(* IEC 61131-3 sources: deprecated-refusr-repo/GP/Main/samples (part 24) *)

(* ---- RND-EXPR_trial-nosed-gunky.st ---- *)
(*
This code implements a randomly grown symbolic expression:

(!(IN26 & (IN45 | ((xor(xor(IN3, !(xor(xor((IN43 & IN34) | (IN19 | IN26), xor(xor(!(IN50), IN21 | IN1), IN17 & IN23)), xor(xor(xor(xor(IN4, IN2), IN41), IN7 & IN29), IN13)))), IN42)) | IN20)))) | (!((xor(xor(!(!(xor(xor(!((!(IN14)) & IN36), ((xor(xor(IN45, IN34), IN41)) | (IN17 | IN11)) & IN16), !(xor(xor(IN37 & IN25, true), IN17 & IN22))))), !((!(IN31)) | (!(IN6)))), ((!(IN16)) | IN27) & (IN46 & ((xor(xor(!(IN15 | IN34), IN28), !(IN7 & IN3))) & ((xor(xor(!(IN32), xor(xor(IN36, IN43), IN28)), !(IN36))) & IN44))))) & IN13))

*)

FUNCTION_BLOCK F_CollectInput
  VAR_IN_OUT
      Data : ARRAY[1..50] OF BOOL;
  END_VAR
  VAR_INPUT
      TICK  : BOOL := 0;
      IN1   : BOOL := 0;
      IN2   : BOOL := 0;
      IN3   : BOOL := 0;
      IN4   : BOOL := 0;
      IN5   : BOOL := 0;
      RESET : BOOL := FALSE;
  END_VAR
  VAR_OUTPUT
      Finished : BOOL;
  END_VAR
  VAR
      j    : USINT := 1;
      tock : BOOL  := 0;
  END_VAR
  IF NOT RESET AND tock = NOT TICK THEN
      Data[j]   := IN1;
      Data[j+1] := IN2;
      Data[j+2] := IN3;
      Data[j+3] := IN4;
      Data[j+4] := IN5;
      j := j + 5;
      tock := TICK;
  ELSE
      j := 1;
      tock := 0;
  END_IF;
  Finished := (j > 50);
END_FUNCTION_BLOCK

PROGRAM Boiler
  VAR
    Data  : ARRAY[1..50] OF BOOL;
    Ready : BOOL;
    CollectInput : F_CollectInput;
  END_VAR
  VAR
    TICK     AT %IX1.0 : BOOL;
    IN1      AT %IX0.3 : BOOL;
    IN2      AT %IX0.4 : BOOL;
    IN3      AT %IX0.5 : BOOL;
    IN4      AT %IX0.6 : BOOL;
    IN5      AT %IX0.7 : BOOL;
    OutReady AT %QX0.0 : BOOL := FALSE;
    FeedNext AT %QX0.1 : BOOL := FALSE;
    Out      AT %QX0.2 : BOOL;
  END_VAR
  CollectInput(TICK:=TICK, IN1:=IN1, IN2:=IN2, IN3:=IN3, IN4:=IN4, IN5:=IN5);
  Ready := CollectInput.Finished;
  FeedNext := 1;
  IF Ready THEN
    Out := ((NOT (Data[26] AND (Data[45] OR (((Data[3] XOR (NOT ((((Data[43] AND Data[34]) OR (Data[19] OR Data[26])) XOR (((NOT Data[50]) XOR (Data[21] OR Data[1])) XOR (Data[17] AND Data[23]))) XOR ((((Data[4] XOR Data[2]) XOR Data[41]) XOR (Data[7] AND Data[29])) XOR Data[13])))) XOR Data[42]) OR Data[20])))) OR (NOT ((((NOT (NOT (((NOT ((NOT Data[14]) AND Data[36])) XOR ((((Data[45] XOR Data[34]) XOR Data[41]) OR (Data[17] OR Data[11])) AND Data[16])) XOR (NOT (((Data[37] AND Data[25]) XOR TRUE) XOR (Data[17] AND Data[22])))))) XOR (NOT ((NOT Data[31]) OR (NOT Data[6])))) XOR (((NOT Data[16]) OR Data[27]) AND (Data[46] AND ((((NOT (Data[15] OR Data[34])) XOR Data[28]) XOR (NOT (Data[7] AND Data[3]))) AND ((((NOT Data[32]) XOR ((Data[36] XOR Data[43]) XOR Data[28])) XOR (NOT Data[36])) AND Data[44]))))) AND Data[13])));
    OutReady := 1;
    CollectInput(RESET:=TRUE);
  END_IF;
END_PROGRAM

CONFIGURATION Config0
  RESOURCE Res0 ON PLC
    TASK task0(INTERVAL := T#20ms,PRIORITY := 0);
    PROGRAM instance0 WITH task0 : Boiler;
  END_RESOURCE
END_CONFIGURATION

(* ---- RND-EXPR_trill-blare-frail.st ---- *)
(*
This code implements a randomly grown symbolic expression:

(xor(xor(xor(xor((((((xor(xor(!(IN12), !(IN17)), xor(xor(IN9, IN18), IN16))) | (!(!(IN37)))) | IN16) & (xor(xor(IN45, (xor(xor(IN41 | IN9, xor(xor(IN35, IN31), IN31)), false & IN31)) | ((xor(xor(IN20, IN44), IN36)) | (IN7 & IN36))), false & IN37))) | IN2) | (IN40 & (xor(xor((xor(xor(xor(xor(IN13, IN26), IN49 | IN33), (xor(xor(IN9, IN4), IN10)) & IN35), (xor(xor(IN38, IN22), IN49)) & (IN26 | IN2))) & (xor(xor((IN21 | IN37) | IN35, xor(xor(xor(xor(IN27, IN35), IN49), IN20), !(IN38))), xor(xor(!(IN24), IN47 & IN9), IN49 & IN17))), (IN2 & ((xor(xor(IN39, true), IN43)) | (!(IN6)))) & (xor(xor(xor(xor(IN32 | IN28, !(IN19)), IN40 | IN22), !(IN3 & IN26)), (IN29 | IN25) | (IN45 & IN27)))), xor(xor((!(IN44)) & IN6, IN29), (!(IN7 & IN11)) | ((false & IN15) | (!(IN19))))))), IN17), xor(xor((IN38 & (IN15 | ((IN27 | (!(IN8))) & (IN23 | (IN11 & IN7))))) | (xor(xor((((xor(xor(IN34, IN2), IN40)) | IN1) | (!(IN9 | IN21))) & (!(xor(xor(IN30 | IN29, xor(xor(IN44, IN42), IN31)), true & IN38))), (IN10 | ((IN10 | IN13) & (IN25 | IN48))) & IN18), xor(xor(!(xor(xor(!(IN15), IN14 & IN49), false)), IN16), IN33))), IN13), xor(xor(!((((!(IN21)) & IN46) | (!(!(IN30)))) | (!((xor(xor(IN29, IN30), IN17)) | (xor(xor(IN48, IN6), IN1))))), xor(xor(!(IN18), (((!(IN34)) & (IN25 | IN49)) & (!(IN46 | IN49))) & (!(xor(xor(xor(xor(IN12, IN43), IN16), IN41), IN17)))), IN11 | (IN5 | false))), ((((!(IN35)) | (xor(xor(IN23, IN39), IN8))) & IN6) & (!(xor(xor(IN21 & IN34, true | IN14), xor(xor(IN23, IN26), IN5))))) & IN28))), !(!(IN4))), (IN38 | (xor(xor(!(IN16 | (IN25 & (!(!(IN31))))), xor(xor(xor(xor((false | (xor(xor(IN33, IN12), IN48))) | ((xor(xor(IN5, IN49), IN14)) & IN11), !((IN49 | IN29) | (IN29 & IN12))), ((IN48 | IN19) | (IN10 | IN4)) | ((!(IN37)) & (IN39 & IN4))), (!((IN33 | true) | (xor(xor(IN26, IN44), IN22)))) | (IN37 | (xor(xor(IN30 | IN33, IN47), !(IN7))))), (!(xor(xor(!(IN21), !(IN11)), !(IN17)))) & IN12)), xor(xor((((!(IN22)) | (IN18 & IN6)) & (xor(xor(xor(xor(IN30, IN18), IN11), IN14 & IN13), IN18 & IN44))) & (xor(xor(IN30 & (IN31 & IN44), xor(xor(xor(xor(IN22, IN16), IN17), xor(xor(IN13, IN42), IN23)), IN38 & IN3)), !(xor(xor(IN41, IN47), IN26)))), IN3), IN12 | IN1)))) & (xor(xor(IN30, !(xor(xor(xor(xor(IN49 & (!(!(IN12))), IN12 & (!(IN13 | IN31))), !((IN21 | IN45) & (IN43 | IN21))), xor(xor(!((IN24 | IN34) | (!(IN1))), ((!(IN44)) & (xor(xor(IN20, IN30), IN17))) | (xor(xor(IN23 & IN49, IN45 & IN25), !(IN34)))), !((!(IN13)) | (xor(xor(IN49, IN15), IN41))))), ((IN4 & (IN19 & IN39)) | ((xor(xor(IN9, IN46), IN40)) & (IN30 & IN45))) & (IN49 | IN13)))), xor(xor(xor(xor(((IN50 & (!(IN24))) & ((IN47 | IN39) & (IN40 & IN24))) & ((xor(xor(IN10 | IN23, IN7 | IN31), IN15 | IN34)) & (IN44 | (!(IN46)))), !(xor(xor(xor(xor(IN29, IN20), IN41 & IN28), IN12), IN27 & (xor(xor(IN42, IN24), IN2))))), IN23), IN11), ((((xor(xor(IN44, IN30), IN46)) | IN35) & IN44) | ((IN45 | (IN7 | IN9)) & IN40)) & IN26))))) | (!((((((xor(xor(IN40, xor(xor(IN25 & IN33, !(IN30)), xor(xor(IN17, IN41), IN29))), IN23)) | (!(xor(xor(xor(xor(IN16, IN49), IN38), IN2 | IN47), IN6 | IN24)))) | IN9) | (!(IN10))) | IN25) & (IN47 | (!(((!(!(IN41 & IN48))) | (IN6 | IN11)) & (((IN12 & IN38) & IN8) | ((xor(xor(IN39 & IN14, IN34 | IN30), xor(xor(IN23, IN46), IN33))) | IN49)))))))

*)

FUNCTION_BLOCK F_CollectInput
  VAR_IN_OUT
      Data : ARRAY[1..50] OF BOOL;
  END_VAR
  VAR_INPUT
      TICK  : BOOL := 0;
      IN1   : BOOL := 0;
      IN2   : BOOL := 0;
      IN3   : BOOL := 0;
      IN4   : BOOL := 0;
      IN5   : BOOL := 0;
      RESET : BOOL := FALSE;
  END_VAR
  VAR_OUTPUT
      Finished : BOOL;
  END_VAR
  VAR
      j    : USINT := 1;
      tock : BOOL  := 0;
  END_VAR
  IF NOT RESET AND tock = NOT TICK THEN
      Data[j]   := IN1;
      Data[j+1] := IN2;
      Data[j+2] := IN3;
      Data[j+3] := IN4;
      Data[j+4] := IN5;
      j := j + 5;
      tock := TICK;
  ELSE
      j := 1;
      tock := 0;
  END_IF;
  Finished := (j > 50);
END_FUNCTION_BLOCK

PROGRAM Boiler
  VAR
    Data  : ARRAY[1..50] OF BOOL;
    Ready : BOOL;
    CollectInput : F_CollectInput;
  END_VAR
  VAR
    TICK     AT %IX1.0 : BOOL;
    IN1      AT %IX0.3 : BOOL;
    IN2      AT %IX0.4 : BOOL;
    IN3      AT %IX0.5 : BOOL;
    IN4      AT %IX0.6 : BOOL;
    IN5      AT %IX0.7 : BOOL;
    OutReady AT %QX0.0 : BOOL := FALSE;
    FeedNext AT %QX0.1 : BOOL := FALSE;
    Out      AT %QX0.2 : BOOL;
  END_VAR
  CollectInput(TICK:=TICK, IN1:=IN1, IN2:=IN2, IN3:=IN3, IN4:=IN4, IN5:=IN5);
  Ready := CollectInput.Finished;
  FeedNext := 1;
  IF Ready THEN
    Out := (((((((((((((NOT Data[12]) XOR (NOT Data[17])) XOR ((Data[9] XOR Data[18]) XOR Data[16])) OR (NOT (NOT Data[37]))) OR Data[16]) AND ((Data[45] XOR ((((Data[41] OR Data[9]) XOR ((Data[35] XOR Data[31]) XOR Data[31])) XOR (FALSE AND Data[31])) OR (((Data[20] XOR Data[44]) XOR Data[36]) OR (Data[7] AND Data[36])))) XOR (FALSE AND Data[37]))) OR Data[2]) OR (Data[40] AND (((((((Data[13] XOR Data[26]) XOR (Data[49] OR Data[33])) XOR (((Data[9] XOR Data[4]) XOR Data[10]) AND Data[35])) XOR (((Data[38] XOR Data[22]) XOR Data[49]) AND (Data[26] OR Data[2]))) AND ((((Data[21] OR Data[37]) OR Data[35]) XOR ((((Data[27] XOR Data[35]) XOR Data[49]) XOR Data[20]) XOR (NOT Data[38]))) XOR (((NOT Data[24]) XOR (Data[47] AND Data[9])) XOR (Data[49] AND Data[17])))) XOR ((Data[2] AND (((Data[39] XOR TRUE) XOR Data[43]) OR (NOT Data[6]))) AND (((((Data[32] OR Data[28]) XOR (NOT Data[19])) XOR (Data[40] OR Data[22])) XOR (NOT (Data[3] AND Data[26]))) XOR ((Data[29] OR Data[25]) OR (Data[45] AND Data[27]))))) XOR ((((NOT Data[44]) AND Data[6]) XOR Data[29]) XOR ((NOT (Data[7] AND Data[11])) OR ((FALSE AND Data[15]) OR (NOT Data[19]))))))) XOR Data[17]) XOR ((((Data[38] AND (Data[15] OR ((Data[27] OR (NOT Data[8])) AND (Data[23] OR (Data[11] AND Data[7]))))) OR (((((((Data[34] XOR Data[2]) XOR Data[40]) OR Data[1]) OR (NOT (Data[9] OR Data[21]))) AND (NOT (((Data[30] OR Data[29]) XOR ((Data[44] XOR Data[42]) XOR Data[31])) XOR (TRUE AND Data[38])))) XOR ((Data[10] OR ((Data[10] OR Data[13]) AND (Data[25] OR Data[48]))) AND Data[18])) XOR (((NOT (((NOT Data[15]) XOR (Data[14] AND Data[49])) XOR FALSE)) XOR Data[16]) XOR Data[33]))) XOR Data[13]) XOR (((NOT ((((NOT Data[21]) AND Data[46]) OR (NOT (NOT Data[30]))) OR (NOT (((Data[29] XOR Data[30]) XOR Data[17]) OR ((Data[48] XOR Data[6]) XOR Data[1]))))) XOR (((NOT Data[18]) XOR ((((NOT Data[34]) AND (Data[25] OR Data[49])) AND (NOT (Data[46] OR Data[49]))) AND (NOT ((((Data[12] XOR Data[43]) XOR Data[16]) XOR Data[41]) XOR Data[17])))) XOR (Data[11] OR (Data[5] OR FALSE)))) XOR (((((NOT Data[35]) OR ((Data[23] XOR Data[39]) XOR Data[8])) AND Data[6]) AND (NOT (((Data[21] AND Data[34]) XOR (TRUE OR Data[14])) XOR ((Data[23] XOR Data[26]) XOR Data[5])))) AND Data[28])))) XOR (NOT (NOT Data[4]))) XOR ((Data[38] OR (((NOT (Data[16] OR (Data[25] AND (NOT (NOT Data[31]))))) XOR ((((((FALSE OR ((Data[33] XOR Data[12]) XOR Data[48])) OR (((Data[5] XOR Data[49]) XOR Data[14]) AND Data[11])) XOR (NOT ((Data[49] OR Data[29]) OR (Data[29] AND Data[12])))) XOR (((Data[48] OR Data[19]) OR (Data[10] OR Data[4])) OR ((NOT Data[37]) AND (Data[39] AND Data[4])))) XOR ((NOT ((Data[33] OR TRUE) OR ((Data[26] XOR Data[44]) XOR Data[22]))) OR (Data[37] OR (((Data[30] OR Data[33]) XOR Data[47]) XOR (NOT Data[7]))))) XOR ((NOT (((NOT Data[21]) XOR (NOT Data[11])) XOR (NOT Data[17]))) AND Data[12]))) XOR ((((((NOT Data[22]) OR (Data[18] AND Data[6])) AND ((((Data[30] XOR Data[18]) XOR Data[11]) XOR (Data[14] AND Data[13])) XOR (Data[18] AND Data[44]))) AND (((Data[30] AND (Data[31] AND Data[44])) XOR ((((Data[22] XOR Data[16]) XOR Data[17]) XOR ((Data[13] XOR Data[42]) XOR Data[23])) XOR (Data[38] AND Data[3]))) XOR (NOT ((Data[41] XOR Data[47]) XOR Data[26])))) XOR Data[3]) XOR (Data[12] OR Data[1])))) AND ((Data[30] XOR (NOT (((((Data[49] AND (NOT (NOT Data[12]))) XOR (Data[12] AND (NOT (Data[13] OR Data[31])))) XOR (NOT ((Data[21] OR Data[45]) AND (Data[43] OR Data[21])))) XOR (((NOT ((Data[24] OR Data[34]) OR (NOT Data[1]))) XOR (((NOT Data[44]) AND ((Data[20] XOR Data[30]) XOR Data[17])) OR (((Data[23] AND Data[49]) XOR (Data[45] AND Data[25])) XOR (NOT Data[34])))) XOR (NOT ((NOT Data[13]) OR ((Data[49] XOR Data[15]) XOR Data[41]))))) XOR (((Data[4] AND (Data[19] AND Data[39])) OR (((Data[9] XOR Data[46]) XOR Data[40]) AND (Data[30] AND Data[45]))) AND (Data[49] OR Data[13]))))) XOR (((((((Data[50] AND (NOT Data[24])) AND ((Data[47] OR Data[39]) AND (Data[40] AND Data[24]))) AND ((((Data[10] OR Data[23]) XOR (Data[7] OR Data[31])) XOR (Data[15] OR Data[34])) AND (Data[44] OR (NOT Data[46])))) XOR (NOT ((((Data[29] XOR Data[20]) XOR (Data[41] AND Data[28])) XOR Data[12]) XOR (Data[27] AND ((Data[42] XOR Data[24]) XOR Data[2]))))) XOR Data[23]) XOR Data[11]) XOR ((((((Data[44] XOR Data[30]) XOR Data[46]) OR Data[35]) AND Data[44]) OR ((Data[45] OR (Data[7] OR Data[9])) AND Data[40])) AND Data[26]))))) OR (NOT (((((((Data[40] XOR (((Data[25] AND Data[33]) XOR (NOT Data[30])) XOR ((Data[17] XOR Data[41]) XOR Data[29]))) XOR Data[23]) OR (NOT ((((Data[16] XOR Data[49]) XOR Data[38]) XOR (Data[2] OR Data[47])) XOR (Data[6] OR Data[24])))) OR Data[9]) OR (NOT Data[10])) OR Data[25]) AND (Data[47] OR (NOT (((NOT (NOT (Data[41] AND Data[48]))) OR (Data[6] OR Data[11])) AND (((Data[12] AND Data[38]) AND Data[8]) OR ((((Data[39] AND Data[14]) XOR (Data[34] OR Data[30])) XOR ((Data[23] XOR Data[46]) XOR Data[33])) OR Data[49]))))))));
    OutReady := 1;
    CollectInput(RESET:=TRUE);
  END_IF;
END_PROGRAM

CONFIGURATION Config0
  RESOURCE Res0 ON PLC
    TASK task0(INTERVAL := T#20ms,PRIORITY := 0);
    PROGRAM instance0 WITH task0 : Boiler;
  END_RESOURCE
END_CONFIGURATION

(* ---- RND-EXPR_tulle-bench-aloha.st ---- *)
(*
This code implements a randomly grown symbolic expression:

(IN29 | (((!(IN27)) | (xor(xor(!(xor(xor(!((!(IN8)) & IN9), xor(xor(xor(xor(xor(xor(IN14, IN9), IN41), xor(xor(IN8, IN28), false)), xor(xor(IN9, IN9), IN2)), !(xor(xor(IN2, IN5), IN41))), (!(IN28)) & (xor(xor(IN12, IN39), IN7)))), IN36)), xor(xor(true, !(((IN30 | IN20) | IN9) & IN3)), xor(xor(false, (!(IN31)) | (xor(xor(IN41 | IN5, IN49 & IN1), !(IN13)))), xor(xor((IN28 | IN50) | (!(IN16)), (xor(xor(IN42, IN4), IN6)) | (xor(xor(IN38, IN42), IN36))), (xor(xor(IN46, IN18), IN35)) & (IN39 & IN11))))), IN39))) & (!(xor(xor(IN22 | ((!(xor(xor(IN21, IN5), IN41 & IN1))) | (xor(xor(xor(xor(IN15 | IN13, IN38 | IN6), !(IN1)), IN29), IN48))), IN18), IN3))))) | (!(!((((IN22 | (xor(xor(!(xor(xor(IN30, false), IN5)), !(IN14 | IN3)), !(IN48)))) | ((((!(IN28)) & (xor(xor(IN29, IN6), IN15))) & ((IN8 & IN49) | IN23)) & (((IN12 & IN1) | (xor(xor(IN43, IN5), IN47))) & ((!(IN33)) | (true | IN20))))) & ((!(IN50 | (!(IN5 | IN30)))) & IN40)) & (xor(xor((xor(xor((xor(xor(xor(xor(IN22, IN30), IN10), IN50), IN23 | IN47)) | (IN1 & (xor(xor(IN46, IN29), IN24))), IN24), ((IN2 & IN18) | (IN26 | IN47)) | ((!(IN19)) & IN35))) | ((IN33 & (!(IN25 | IN20))) | (xor(xor((xor(xor(IN40, IN13), IN19)) & (xor(xor(IN2, IN37), IN10)), (IN49 | IN40) & IN19), (xor(xor(IN25, IN24), IN14)) & (IN22 & IN32)))), (!(!((xor(xor(IN42, IN8), IN1)) & (!(IN42))))) & ((!(IN23 & IN19)) | ((!(IN29 & IN50)) & (!(IN8 & IN35))))), !(xor(xor(xor(xor((IN29 & IN22) & (!(IN14)), (IN32 & IN20) & (xor(xor(IN7, IN24), IN7))), (true & IN45) | (IN31 | IN44)), (xor(xor(!(IN45), IN35 | IN9), IN40 | IN3)) | ((xor(xor(IN5, IN37), IN27)) | (xor(xor(IN25, IN45), IN32)))), (false & (IN9 | IN18)) | (xor(xor(IN8, xor(xor(IN10, IN26), IN25)), !(IN39))))))))))

*)

FUNCTION_BLOCK F_CollectInput
  VAR_IN_OUT
      Data : ARRAY[1..50] OF BOOL;
  END_VAR
  VAR_INPUT
      TICK  : BOOL := 0;
      IN1   : BOOL := 0;
      IN2   : BOOL := 0;
      IN3   : BOOL := 0;
      IN4   : BOOL := 0;
      IN5   : BOOL := 0;
      RESET : BOOL := FALSE;
  END_VAR
  VAR_OUTPUT
      Finished : BOOL;
  END_VAR
  VAR
      j    : USINT := 1;
      tock : BOOL  := 0;
  END_VAR
  IF NOT RESET AND tock = NOT TICK THEN
      Data[j]   := IN1;
      Data[j+1] := IN2;
      Data[j+2] := IN3;
      Data[j+3] := IN4;
      Data[j+4] := IN5;
      j := j + 5;
      tock := TICK;
  ELSE
      j := 1;
      tock := 0;
  END_IF;
  Finished := (j > 50);
END_FUNCTION_BLOCK

PROGRAM Boiler
  VAR
    Data  : ARRAY[1..50] OF BOOL;
    Ready : BOOL;
    CollectInput : F_CollectInput;
  END_VAR
  VAR
    TICK     AT %IX1.0 : BOOL;
    IN1      AT %IX0.3 : BOOL;
    IN2      AT %IX0.4 : BOOL;
    IN3      AT %IX0.5 : BOOL;
    IN4      AT %IX0.6 : BOOL;
    IN5      AT %IX0.7 : BOOL;
    OutReady AT %QX0.0 : BOOL := FALSE;
    FeedNext AT %QX0.1 : BOOL := FALSE;
    Out      AT %QX0.2 : BOOL;
  END_VAR
  CollectInput(TICK:=TICK, IN1:=IN1, IN2:=IN2, IN3:=IN3, IN4:=IN4, IN5:=IN5);
  Ready := CollectInput.Finished;
  FeedNext := 1;
  IF Ready THEN
    Out := ((Data[29] OR (((NOT Data[27]) OR (((NOT (((NOT ((NOT Data[8]) AND Data[9])) XOR ((((((Data[14] XOR Data[9]) XOR Data[41]) XOR ((Data[8] XOR Data[28]) XOR FALSE)) XOR ((Data[9] XOR Data[9]) XOR Data[2])) XOR (NOT ((Data[2] XOR Data[5]) XOR Data[41]))) XOR ((NOT Data[28]) AND ((Data[12] XOR Data[39]) XOR Data[7])))) XOR Data[36])) XOR ((TRUE XOR (NOT (((Data[30] OR Data[20]) OR Data[9]) AND Data[3]))) XOR ((FALSE XOR ((NOT Data[31]) OR (((Data[41] OR Data[5]) XOR (Data[49] AND Data[1])) XOR (NOT Data[13])))) XOR ((((Data[28] OR Data[50]) OR (NOT Data[16])) XOR (((Data[42] XOR Data[4]) XOR Data[6]) OR ((Data[38] XOR Data[42]) XOR Data[36]))) XOR (((Data[46] XOR Data[18]) XOR Data[35]) AND (Data[39] AND Data[11])))))) XOR Data[39])) AND (NOT (((Data[22] OR ((NOT ((Data[21] XOR Data[5]) XOR (Data[41] AND Data[1]))) OR (((((Data[15] OR Data[13]) XOR (Data[38] OR Data[6])) XOR (NOT Data[1])) XOR Data[29]) XOR Data[48]))) XOR Data[18]) XOR Data[3])))) OR (NOT (NOT ((((Data[22] OR (((NOT ((Data[30] XOR FALSE) XOR Data[5])) XOR (NOT (Data[14] OR Data[3]))) XOR (NOT Data[48]))) OR ((((NOT Data[28]) AND ((Data[29] XOR Data[6]) XOR Data[15])) AND ((Data[8] AND Data[49]) OR Data[23])) AND (((Data[12] AND Data[1]) OR ((Data[43] XOR Data[5]) XOR Data[47])) AND ((NOT Data[33]) OR (TRUE OR Data[20]))))) AND ((NOT (Data[50] OR (NOT (Data[5] OR Data[30])))) AND Data[40])) AND ((((((((((Data[22] XOR Data[30]) XOR Data[10]) XOR Data[50]) XOR (Data[23] OR Data[47])) OR (Data[1] AND ((Data[46] XOR Data[29]) XOR Data[24]))) XOR Data[24]) XOR (((Data[2] AND Data[18]) OR (Data[26] OR Data[47])) OR ((NOT Data[19]) AND Data[35]))) OR ((Data[33] AND (NOT (Data[25] OR Data[20]))) OR (((((Data[40] XOR Data[13]) XOR Data[19]) AND ((Data[2] XOR Data[37]) XOR Data[10])) XOR ((Data[49] OR Data[40]) AND Data[19])) XOR (((Data[25] XOR Data[24]) XOR Data[14]) AND (Data[22] AND Data[32]))))) XOR ((NOT (NOT (((Data[42] XOR Data[8]) XOR Data[1]) AND (NOT Data[42])))) AND ((NOT (Data[23] AND Data[19])) OR ((NOT (Data[29] AND Data[50])) AND (NOT (Data[8] AND Data[35])))))) XOR (NOT ((((((Data[29] AND Data[22]) AND (NOT Data[14])) XOR ((Data[32] AND Data[20]) AND ((Data[7] XOR Data[24]) XOR Data[7]))) XOR ((TRUE AND Data[45]) OR (Data[31] OR Data[44]))) XOR ((((NOT Data[45]) XOR (Data[35] OR Data[9])) XOR (Data[40] OR Data[3])) OR (((Data[5] XOR Data[37]) XOR Data[27]) OR ((Data[25] XOR Data[45]) XOR Data[32])))) XOR ((FALSE AND (Data[9] OR Data[18])) OR ((Data[8] XOR ((Data[10] XOR Data[26]) XOR Data[25])) XOR (NOT Data[39]))))))))));
    OutReady := 1;
    CollectInput(RESET:=TRUE);
  END_IF;
END_PROGRAM

CONFIGURATION Config0
  RESOURCE Res0 ON PLC
    TASK task0(INTERVAL := T#20ms,PRIORITY := 0);
    PROGRAM instance0 WITH task0 : Boiler;
  END_RESOURCE
END_CONFIGURATION

(* ---- RND-EXPR_umped-hades-orlon.st ---- *)
(*
This code implements a randomly grown symbolic expression:

xor(xor(!((!(((xor(xor(((!(IN45)) & (IN32 | IN40)) & ((IN23 | IN38) | (!(IN24))), xor(xor((IN15 | IN19) & IN39, !(IN4 & IN13)), (xor(xor(IN43, IN11), IN25)) & (IN25 | IN49))), IN19)) | (xor(xor(IN43 & ((IN16 & IN26) | (!(IN43))), IN24 | ((!(IN13)) | IN33)), xor(xor(IN32, (IN20 & IN40) | (IN18 | IN23)), (IN42 & IN39) & (!(IN6)))))) & (!(IN16 & (xor(xor(!(IN50 & IN37), IN25), IN4)))))) & (!(!(((!(xor(xor(IN29 | IN47, xor(xor(IN44, IN42), IN1)), IN48 & IN20))) & (xor(xor((!(IN19)) | (IN47 & IN15), !(xor(xor(IN3, IN39), IN10))), xor(xor(IN35, IN48), IN40 & IN6)))) | (xor(xor(IN2, IN12), !(IN1))))))), IN30 | ((((xor(xor(((xor(xor(IN20 & IN48, !(IN20)), xor(xor(IN21, IN15), IN38))) & ((!(IN47)) & (IN13 & IN31))) & IN25, (((!(IN17)) | (IN34 | IN40)) | IN35) | ((xor(xor(IN37 | IN35, IN11 | IN33), !(IN9))) & ((IN43 & IN14) & (!(IN26))))), (xor(xor(xor(xor(IN45 & IN37, !(IN12)), IN4 | IN33), xor(xor(IN40, IN6 | IN14), IN38)), xor(xor(IN47 & IN30, IN29), !(IN36)))) | ((!(IN17)) | (xor(xor(IN45 | IN20, IN46 & IN36), !(IN17)))))) & (IN31 | (!(((IN9 | IN39) | (IN1 | IN44)) | (!(IN39 | IN42)))))) & IN41) & (((xor(xor(!(IN41 & (xor(xor(IN26 | IN47, xor(xor(IN25, IN44), IN28)), !(IN22)))), IN30), !(!(IN7 | (xor(xor(IN15, IN18), IN35)))))) | IN43) & (((xor(xor((xor(xor(!(IN37), xor(xor(IN36, IN29), IN20)), IN45)) | (xor(xor(IN24, xor(xor(IN17, IN22), IN40)), IN33 & IN36)), xor(xor(IN9 & (xor(xor(IN8, IN7), IN1)), IN29 | (IN49 | IN38)), xor(xor(IN48 | IN37, xor(xor(IN40, IN21), IN27)), !(IN9)))), !((xor(xor(IN21, IN35), IN17)) | IN47))) | IN41) | (IN40 & ((!(xor(xor(IN14 | IN35, IN10), true & IN31))) & (xor(xor((!(IN11)) | (!(IN1)), IN28), xor(xor(IN12, IN14 | IN38), IN26 & IN23))))))))), false)

*)

FUNCTION_BLOCK F_CollectInput
  VAR_IN_OUT
      Data : ARRAY[1..50] OF BOOL;
  END_VAR
  VAR_INPUT
      TICK  : BOOL := 0;
      IN1   : BOOL := 0;
      IN2   : BOOL := 0;
      IN3   : BOOL := 0;
      IN4   : BOOL := 0;
      IN5   : BOOL := 0;
      RESET : BOOL := FALSE;
  END_VAR
  VAR_OUTPUT
      Finished : BOOL;
  END_VAR
  VAR
      j    : USINT := 1;
      tock : BOOL  := 0;
  END_VAR
  IF NOT RESET AND tock = NOT TICK THEN
      Data[j]   := IN1;
      Data[j+1] := IN2;
      Data[j+2] := IN3;
      Data[j+3] := IN4;
      Data[j+4] := IN5;
      j := j + 5;
      tock := TICK;
  ELSE
      j := 1;
      tock := 0;
  END_IF;
  Finished := (j > 50);
END_FUNCTION_BLOCK

PROGRAM Boiler
  VAR
    Data  : ARRAY[1..50] OF BOOL;
    Ready : BOOL;
    CollectInput : F_CollectInput;
  END_VAR
  VAR
    TICK     AT %IX1.0 : BOOL;
    IN1      AT %IX0.3 : BOOL;
    IN2      AT %IX0.4 : BOOL;
    IN3      AT %IX0.5 : BOOL;
    IN4      AT %IX0.6 : BOOL;
    IN5      AT %IX0.7 : BOOL;
    OutReady AT %QX0.0 : BOOL := FALSE;
    FeedNext AT %QX0.1 : BOOL := FALSE;
    Out      AT %QX0.2 : BOOL;
  END_VAR
  CollectInput(TICK:=TICK, IN1:=IN1, IN2:=IN2, IN3:=IN3, IN4:=IN4, IN5:=IN5);
  Ready := CollectInput.Finished;
  FeedNext := 1;
  IF Ready THEN
    Out := (((NOT ((NOT (((((((NOT Data[45]) AND (Data[32] OR Data[40])) AND ((Data[23] OR Data[38]) OR (NOT Data[24]))) XOR ((((Data[15] OR Data[19]) AND Data[39]) XOR (NOT (Data[4] AND Data[13]))) XOR (((Data[43] XOR Data[11]) XOR Data[25]) AND (Data[25] OR Data[49])))) XOR Data[19]) OR (((Data[43] AND ((Data[16] AND Data[26]) OR (NOT Data[43]))) XOR (Data[24] OR ((NOT Data[13]) OR Data[33]))) XOR ((Data[32] XOR ((Data[20] AND Data[40]) OR (Data[18] OR Data[23]))) XOR ((Data[42] AND Data[39]) AND (NOT Data[6]))))) AND (NOT (Data[16] AND (((NOT (Data[50] AND Data[37])) XOR Data[25]) XOR Data[4]))))) AND (NOT (NOT (((NOT (((Data[29] OR Data[47]) XOR ((Data[44] XOR Data[42]) XOR Data[1])) XOR (Data[48] AND Data[20]))) AND ((((NOT Data[19]) OR (Data[47] AND Data[15])) XOR (NOT ((Data[3] XOR Data[39]) XOR Data[10]))) XOR ((Data[35] XOR Data[48]) XOR (Data[40] AND Data[6])))) OR ((Data[2] XOR Data[12]) XOR (NOT Data[1]))))))) XOR (Data[30] OR ((((((((((Data[20] AND Data[48]) XOR (NOT Data[20])) XOR ((Data[21] XOR Data[15]) XOR Data[38])) AND ((NOT Data[47]) AND (Data[13] AND Data[31]))) AND Data[25]) XOR ((((NOT Data[17]) OR (Data[34] OR Data[40])) OR Data[35]) OR ((((Data[37] OR Data[35]) XOR (Data[11] OR Data[33])) XOR (NOT Data[9])) AND ((Data[43] AND Data[14]) AND (NOT Data[26]))))) XOR ((((((Data[45] AND Data[37]) XOR (NOT Data[12])) XOR (Data[4] OR Data[33])) XOR ((Data[40] XOR (Data[6] OR Data[14])) XOR Data[38])) XOR (((Data[47] AND Data[30]) XOR Data[29]) XOR (NOT Data[36]))) OR ((NOT Data[17]) OR (((Data[45] OR Data[20]) XOR (Data[46] AND Data[36])) XOR (NOT Data[17]))))) AND (Data[31] OR (NOT (((Data[9] OR Data[39]) OR (Data[1] OR Data[44])) OR (NOT (Data[39] OR Data[42])))))) AND Data[41]) AND (((((NOT (Data[41] AND (((Data[26] OR Data[47]) XOR ((Data[25] XOR Data[44]) XOR Data[28])) XOR (NOT Data[22])))) XOR Data[30]) XOR (NOT (NOT (Data[7] OR ((Data[15] XOR Data[18]) XOR Data[35]))))) OR Data[43]) AND ((((((((NOT Data[37]) XOR ((Data[36] XOR Data[29]) XOR Data[20])) XOR Data[45]) OR ((Data[24] XOR ((Data[17] XOR Data[22]) XOR Data[40])) XOR (Data[33] AND Data[36]))) XOR (((Data[9] AND ((Data[8] XOR Data[7]) XOR Data[1])) XOR (Data[29] OR (Data[49] OR Data[38]))) XOR (((Data[48] OR Data[37]) XOR ((Data[40] XOR Data[21]) XOR Data[27])) XOR (NOT Data[9])))) XOR (NOT (((Data[21] XOR Data[35]) XOR Data[17]) OR Data[47]))) OR Data[41]) OR (Data[40] AND ((NOT (((Data[14] OR Data[35]) XOR Data[10]) XOR (TRUE AND Data[31]))) AND ((((NOT Data[11]) OR (NOT Data[1])) XOR Data[28]) XOR ((Data[12] XOR (Data[14] OR Data[38])) XOR (Data[26] AND Data[23])))))))))) XOR FALSE);
    OutReady := 1;
    CollectInput(RESET:=TRUE);
  END_IF;
END_PROGRAM

CONFIGURATION Config0
  RESOURCE Res0 ON PLC
    TASK task0(INTERVAL := T#20ms,PRIORITY := 0);
    PROGRAM instance0 WITH task0 : Boiler;
  END_RESOURCE
END_CONFIGURATION

(* ---- RND-EXPR_unapt-filch-drawn.st ---- *)
(*
This code implements a randomly grown symbolic expression:

(!(((xor(xor(((xor(xor((xor(xor(IN31, IN18), IN21)) & (IN50 & IN24), IN29), xor(xor(IN25, IN42 | IN8), !(IN3)))) & IN26) & IN17, xor(xor((!((xor(xor(IN20, IN38), IN31)) | (xor(xor(IN29, IN48), IN28)))) | (!((!(IN37)) | (IN38 & IN28))), xor(xor(xor(xor((xor(xor(IN30, IN11), IN47)) & (IN32 | IN44), IN25), (xor(xor(IN31, IN27), IN19)) | (xor(xor(IN40, IN1), IN7))), xor(xor((IN42 | IN13) & IN35, IN34), IN17)), IN21)), xor(xor(IN8, !(IN18)), (IN32 | (xor(xor(IN10, IN41), IN41))) | ((!(IN50)) & (IN29 & true))))), IN27)) | ((xor(xor(!((xor(xor(IN22 | IN34, !(IN37)), xor(xor(IN11, IN3), IN46))) & ((!(IN45)) & (IN17 | IN31))), (xor(xor(IN6, xor(xor(IN43 & IN8, IN41 | IN39), xor(xor(IN17, IN48), IN34))), !(IN3 & IN25))) | (!((IN48 | IN11) & (IN44 & IN29)))), (xor(xor(IN34, IN28), IN1)) | ((xor(xor(IN10 | IN34, IN26 & IN10), xor(xor(IN27, IN4), IN46))) & true))) & (xor(xor(IN9 | (((!(IN18)) | (IN7 | IN8)) | (xor(xor(IN40 & IN19, IN19), IN7 | IN35))), xor(xor(IN17 | (xor(xor(IN9 | IN10, IN25 | IN22), IN44 & IN10)), !(IN31)), ((xor(xor(IN43, IN15), IN11)) & (IN26 & IN1)) & (!(!(IN17))))), IN36)))) & ((xor(xor(!(xor(xor((xor(xor(IN32 | IN14, IN28), IN24 | IN36)) & ((!(IN49)) & IN22), ((!(IN46)) | (xor(xor(IN24, IN40), IN38))) & (xor(xor(IN3, !(IN41)), IN31))), IN18 & ((xor(xor(IN34, IN9), IN47)) & IN21))), !(xor(xor(((xor(xor(IN16, false), IN31)) | (IN27 & IN33)) & ((IN22 & IN17) & IN46), xor(xor(!(IN36 | IN48), !(IN9)), (!(IN16)) | IN39)), (xor(xor(IN14 & IN26, !(IN31)), !(IN12))) | ((IN9 | IN16) | (IN37 & IN9))))), ((xor(xor(xor(xor(IN11, IN9 & IN18), xor(xor(IN9, IN14), IN5)), (IN32 & IN47) & (xor(xor(IN18, IN46), IN41))), (xor(xor(IN45, IN26), IN7)) & (xor(xor(IN40, IN29), IN50)))) & (!(IN37 & (IN48 & IN30)))) | ((!((!(IN43)) & (IN30 | IN26))) | ((!(IN22 & IN10)) & ((xor(xor(IN22, IN47), IN12)) | IN24))))) & (xor(xor(IN49, (!(!(xor(xor(IN8 & IN39, xor(xor(IN12, IN8), IN5)), IN14 & IN35)))) & (((!(IN16 | IN46)) | IN18) | IN36)), !((xor(xor((xor(xor(IN23, IN13), IN21)) & (!(IN19)), (!(IN36)) & (IN14 & IN28)), (xor(xor(true, IN35), IN6)) & (IN19 & IN14))) | (xor(xor((xor(xor(IN22, IN43), IN42)) | (!(IN39)), IN43), (IN8 & IN30) | IN2)))))))) | (!((xor(xor(((!(xor(xor((IN27 & IN6) | (IN50 | IN7), false), xor(xor(!(IN35), IN6 | IN35), IN48 | IN2)))) & (!(!((IN2 | IN21) & (IN26 & IN21))))) & (!(!(!(IN29)))), IN19 | IN3), !((xor(xor(!((IN49 & true) | (IN42 | IN48)), (!(xor(xor(IN44, IN22), IN44))) & (!(IN9 & IN13))), IN1)) | (((xor(xor(IN11, xor(xor(IN23, IN30), IN25)), IN39 & IN10)) & (!(!(IN33)))) | (((!(IN24)) | (!(IN39))) | true))))) | ((!((xor(xor((!(!(IN14))) | IN12, !((!(IN1)) & (!(IN37)))), xor(xor(xor(xor(IN4, IN1 & IN46), IN26), xor(xor(true, IN13 | IN15), IN21 & IN49)), !(IN41 & IN44)))) | ((!(false | (IN2 & IN14))) & (((IN15 & IN28) | (xor(xor(IN6, IN46), IN18))) & (xor(xor(IN5 | IN17, xor(xor(IN11, IN36), IN45)), IN43)))))) | (xor(xor(IN37, !(xor(xor((IN33 & IN26) & (xor(xor(xor(xor(IN24, IN11), IN28), !(IN46)), IN24 & IN37)), IN2), xor(xor(!(IN50), (xor(xor(IN43, IN46), IN48)) & (IN11 & IN26)), (!(IN45)) & (!(IN37)))))), (xor(xor(IN37, (xor(xor(IN2 | IN8, IN15), IN33 & IN32)) | (!(IN23 | false))), (!(IN15 | IN3)) & (xor(xor(IN22, IN46), !(IN26))))) & (IN43 | IN25))))))

*)

FUNCTION_BLOCK F_CollectInput
  VAR_IN_OUT
      Data : ARRAY[1..50] OF BOOL;
  END_VAR
  VAR_INPUT
      TICK  : BOOL := 0;
      IN1   : BOOL := 0;
      IN2   : BOOL := 0;
      IN3   : BOOL := 0;
      IN4   : BOOL := 0;
      IN5   : BOOL := 0;
      RESET : BOOL := FALSE;
  END_VAR
  VAR_OUTPUT
      Finished : BOOL;
  END_VAR
  VAR
      j    : USINT := 1;
      tock : BOOL  := 0;
  END_VAR
  IF NOT RESET AND tock = NOT TICK THEN
      Data[j]   := IN1;
      Data[j+1] := IN2;
      Data[j+2] := IN3;
      Data[j+3] := IN4;
      Data[j+4] := IN5;
      j := j + 5;
      tock := TICK;
  ELSE
      j := 1;
      tock := 0;
  END_IF;
  Finished := (j > 50);
END_FUNCTION_BLOCK

PROGRAM Boiler
  VAR
    Data  : ARRAY[1..50] OF BOOL;
    Ready : BOOL;
    CollectInput : F_CollectInput;
  END_VAR
  VAR
    TICK     AT %IX1.0 : BOOL;
    IN1      AT %IX0.3 : BOOL;
    IN2      AT %IX0.4 : BOOL;
    IN3      AT %IX0.5 : BOOL;
    IN4      AT %IX0.6 : BOOL;
    IN5      AT %IX0.7 : BOOL;
    OutReady AT %QX0.0 : BOOL := FALSE;
    FeedNext AT %QX0.1 : BOOL := FALSE;
    Out      AT %QX0.2 : BOOL;
  END_VAR
  CollectInput(TICK:=TICK, IN1:=IN1, IN2:=IN2, IN3:=IN3, IN4:=IN4, IN5:=IN5);
  Ready := CollectInput.Finished;
  FeedNext := 1;
  IF Ready THEN
    Out := ((NOT (((((((((((Data[31] XOR Data[18]) XOR Data[21]) AND (Data[50] AND Data[24])) XOR Data[29]) XOR ((Data[25] XOR (Data[42] OR Data[8])) XOR (NOT Data[3]))) AND Data[26]) AND Data[17]) XOR ((((NOT (((Data[20] XOR Data[38]) XOR Data[31]) OR ((Data[29] XOR Data[48]) XOR Data[28]))) OR (NOT ((NOT Data[37]) OR (Data[38] AND Data[28])))) XOR (((((((Data[30] XOR Data[11]) XOR Data[47]) AND (Data[32] OR Data[44])) XOR Data[25]) XOR (((Data[31] XOR Data[27]) XOR Data[19]) OR ((Data[40] XOR Data[1]) XOR Data[7]))) XOR ((((Data[42] OR Data[13]) AND Data[35]) XOR Data[34]) XOR Data[17])) XOR Data[21])) XOR ((Data[8] XOR (NOT Data[18])) XOR ((Data[32] OR ((Data[10] XOR Data[41]) XOR Data[41])) OR ((NOT Data[50]) AND (Data[29] AND TRUE)))))) XOR Data[27]) OR ((((NOT ((((Data[22] OR Data[34]) XOR (NOT Data[37])) XOR ((Data[11] XOR Data[3]) XOR Data[46])) AND ((NOT Data[45]) AND (Data[17] OR Data[31])))) XOR (((Data[6] XOR (((Data[43] AND Data[8]) XOR (Data[41] OR Data[39])) XOR ((Data[17] XOR Data[48]) XOR Data[34]))) XOR (NOT (Data[3] AND Data[25]))) OR (NOT ((Data[48] OR Data[11]) AND (Data[44] AND Data[29]))))) XOR (((Data[34] XOR Data[28]) XOR Data[1]) OR ((((Data[10] OR Data[34]) XOR (Data[26] AND Data[10])) XOR ((Data[27] XOR Data[4]) XOR Data[46])) AND TRUE))) AND (((Data[9] OR (((NOT Data[18]) OR (Data[7] OR Data[8])) OR (((Data[40] AND Data[19]) XOR Data[19]) XOR (Data[7] OR Data[35])))) XOR (((Data[17] OR (((Data[9] OR Data[10]) XOR (Data[25] OR Data[22])) XOR (Data[44] AND Data[10]))) XOR (NOT Data[31])) XOR ((((Data[43] XOR Data[15]) XOR Data[11]) AND (Data[26] AND Data[1])) AND (NOT (NOT Data[17]))))) XOR Data[36]))) AND ((((NOT ((((((Data[32] OR Data[14]) XOR Data[28]) XOR (Data[24] OR Data[36])) AND ((NOT Data[49]) AND Data[22])) XOR (((NOT Data[46]) OR ((Data[24] XOR Data[40]) XOR Data[38])) AND ((Data[3] XOR (NOT Data[41])) XOR Data[31]))) XOR (Data[18] AND (((Data[34] XOR Data[9]) XOR Data[47]) AND Data[21])))) XOR (NOT ((((((Data[16] XOR FALSE) XOR Data[31]) OR (Data[27] AND Data[33])) AND ((Data[22] AND Data[17]) AND Data[46])) XOR (((NOT (Data[36] OR Data[48])) XOR (NOT Data[9])) XOR ((NOT Data[16]) OR Data[39]))) XOR ((((Data[14] AND Data[26]) XOR (NOT Data[31])) XOR (NOT Data[12])) OR ((Data[9] OR Data[16]) OR (Data[37] AND Data[9])))))) XOR ((((((Data[11] XOR (Data[9] AND Data[18])) XOR ((Data[9] XOR Data[14]) XOR Data[5])) XOR ((Data[32] AND Data[47]) AND ((Data[18] XOR Data[46]) XOR Data[41]))) XOR (((Data[45] XOR Data[26]) XOR Data[7]) AND ((Data[40] XOR Data[29]) XOR Data[50]))) AND (NOT (Data[37] AND (Data[48] AND Data[30])))) OR ((NOT ((NOT Data[43]) AND (Data[30] OR Data[26]))) OR ((NOT (Data[22] AND Data[10])) AND (((Data[22] XOR Data[47]) XOR Data[12]) OR Data[24]))))) AND ((Data[49] XOR ((NOT (NOT (((Data[8] AND Data[39]) XOR ((Data[12] XOR Data[8]) XOR Data[5])) XOR (Data[14] AND Data[35])))) AND (((NOT (Data[16] OR Data[46])) OR Data[18]) OR Data[36]))) XOR (NOT ((((((Data[23] XOR Data[13]) XOR Data[21]) AND (NOT Data[19])) XOR ((NOT Data[36]) AND (Data[14] AND Data[28]))) XOR (((TRUE XOR Data[35]) XOR Data[6]) AND (Data[19] AND Data[14]))) OR (((((Data[22] XOR Data[43]) XOR Data[42]) OR (NOT Data[39])) XOR Data[43]) XOR ((Data[8] AND Data[30]) OR Data[2])))))))) OR (NOT ((((((NOT ((((Data[27] AND Data[6]) OR (Data[50] OR Data[7])) XOR FALSE) XOR (((NOT Data[35]) XOR (Data[6] OR Data[35])) XOR (Data[48] OR Data[2])))) AND (NOT (NOT ((Data[2] OR Data[21]) AND (Data[26] AND Data[21]))))) AND (NOT (NOT (NOT Data[29])))) XOR (Data[19] OR Data[3])) XOR (NOT ((((NOT ((Data[49] AND TRUE) OR (Data[42] OR Data[48]))) XOR ((NOT ((Data[44] XOR Data[22]) XOR Data[44])) AND (NOT (Data[9] AND Data[13])))) XOR Data[1]) OR ((((Data[11] XOR ((Data[23] XOR Data[30]) XOR Data[25])) XOR (Data[39] AND Data[10])) AND (NOT (NOT Data[33]))) OR (((NOT Data[24]) OR (NOT Data[39])) OR TRUE))))) OR ((NOT (((((NOT (NOT Data[14])) OR Data[12]) XOR (NOT ((NOT Data[1]) AND (NOT Data[37])))) XOR ((((Data[4] XOR (Data[1] AND Data[46])) XOR Data[26]) XOR ((TRUE XOR (Data[13] OR Data[15])) XOR (Data[21] AND Data[49]))) XOR (NOT (Data[41] AND Data[44])))) OR ((NOT (FALSE OR (Data[2] AND Data[14]))) AND (((Data[15] AND Data[28]) OR ((Data[6] XOR Data[46]) XOR Data[18])) AND (((Data[5] OR Data[17]) XOR ((Data[11] XOR Data[36]) XOR Data[45])) XOR Data[43]))))) OR ((Data[37] XOR (NOT ((((Data[33] AND Data[26]) AND ((((Data[24] XOR Data[11]) XOR Data[28]) XOR (NOT Data[46])) XOR (Data[24] AND Data[37]))) XOR Data[2]) XOR (((NOT Data[50]) XOR (((Data[43] XOR Data[46]) XOR Data[48]) AND (Data[11] AND Data[26]))) XOR ((NOT Data[45]) AND (NOT Data[37])))))) XOR (((Data[37] XOR ((((Data[2] OR Data[8]) XOR Data[15]) XOR (Data[33] AND Data[32])) OR (NOT (Data[23] OR FALSE)))) XOR ((NOT (Data[15] OR Data[3])) AND ((Data[22] XOR Data[46]) XOR (NOT Data[26])))) AND (Data[43] OR Data[25])))))));
    OutReady := 1;
    CollectInput(RESET:=TRUE);
  END_IF;
END_PROGRAM

CONFIGURATION Config0
  RESOURCE Res0 ON PLC
    TASK task0(INTERVAL := T#20ms,PRIORITY := 0);
    PROGRAM instance0 WITH task0 : Boiler;
  END_RESOURCE
END_CONFIGURATION

(* ---- RND-EXPR_undid-rasps-zebra.st ---- *)
(*
This code implements a randomly grown symbolic expression:

(!(IN26)) & (xor(xor(!(IN23), !(!((((xor(xor((!(IN29)) | (!(IN21)), xor(xor(xor(xor(true, IN46), IN14), !(IN7)), !(IN19))), !(IN12))) & ((!(!(IN9))) | IN10)) | (!(IN29 & IN6))) & ((xor(xor(IN34, IN46), !((IN47 | IN39) & (xor(xor(IN48, IN16), IN35))))) | (xor(xor(xor(xor(xor(xor(IN18, !(IN46)), IN4), false & (!(IN20))), !(!(IN26))), false), IN34 | (xor(xor(xor(xor(IN48, IN50), IN49), !(IN38)), IN45 & IN13)))))))), (xor(xor((!((!(xor(xor(false, !(IN30)), IN27))) | (xor(xor(xor(xor(IN25 & IN4, IN3 | IN3), IN47 & IN26), !(IN25 & IN25)), !(!(IN24)))))) | (((!(IN21 | (IN5 & IN39))) & ((xor(xor(IN3 & IN24, IN49 & IN44), IN24 & IN39)) | ((IN21 | IN27) & IN42))) & (xor(xor(((!(IN46)) & (xor(xor(IN42, IN44), IN38))) & false, xor(xor(xor(xor(IN38 & false, IN32), !(IN21)), (xor(xor(IN22, IN10), IN42)) & (false | IN15)), IN12)), xor(xor(IN22 | (IN41 | IN39), (IN23 | IN41) & (IN23 & IN21)), (!(IN22)) | (xor(xor(IN47, IN35), IN37)))))), xor(xor(!((((IN13 & IN38) | (!(IN21))) | IN42) | (((IN34 & IN31) | (IN6 & IN28)) | ((IN45 & IN33) | IN42))), xor(xor(IN1, (((IN32 & IN43) & (IN10 | IN49)) & (xor(xor(xor(xor(IN42, IN8), IN40), IN12 | IN31), IN25 & IN30))) | IN13), xor(xor(xor(xor(false & (IN14 & IN9), !(IN3)), IN39 & (IN11 & IN35)), IN27 | (!(IN6 | IN39))), !(xor(xor(!(IN37), xor(xor(IN1, IN13), IN25)), xor(xor(IN22, false), IN17)))))), IN31 | (xor(xor(((!(IN11)) & (xor(xor(IN10, IN29), IN38))) | ((IN20 & IN29) | (!(IN22))), IN19), xor(xor((IN1 | IN39) | IN22, (!(IN7)) & (IN26 | IN10)), IN12))))), !(xor(xor(!(IN9), ((IN38 & (!(IN35))) & (!(IN32 | IN20))) & (xor(xor(true, xor(xor(IN35, IN33 | IN35), IN10 | IN17)), IN42 & (xor(xor(IN28, IN5), IN11))))), IN27 & (IN1 | ((!(IN45)) & (IN8 & IN17))))))) | (!(!(IN22)))))

*)

FUNCTION_BLOCK F_CollectInput
  VAR_IN_OUT
      Data : ARRAY[1..50] OF BOOL;
  END_VAR
  VAR_INPUT
      TICK  : BOOL := 0;
      IN1   : BOOL := 0;
      IN2   : BOOL := 0;
      IN3   : BOOL := 0;
      IN4   : BOOL := 0;
      IN5   : BOOL := 0;
      RESET : BOOL := FALSE;
  END_VAR
  VAR_OUTPUT
      Finished : BOOL;
  END_VAR
  VAR
      j    : USINT := 1;
      tock : BOOL  := 0;
  END_VAR
  IF NOT RESET AND tock = NOT TICK THEN
      Data[j]   := IN1;
      Data[j+1] := IN2;
      Data[j+2] := IN3;
      Data[j+3] := IN4;
      Data[j+4] := IN5;
      j := j + 5;
      tock := TICK;
  ELSE
      j := 1;
      tock := 0;
  END_IF;
  Finished := (j > 50);
END_FUNCTION_BLOCK

PROGRAM Boiler
  VAR
    Data  : ARRAY[1..50] OF BOOL;
    Ready : BOOL;
    CollectInput : F_CollectInput;
  END_VAR
  VAR
    TICK     AT %IX1.0 : BOOL;
    IN1      AT %IX0.3 : BOOL;
    IN2      AT %IX0.4 : BOOL;
    IN3      AT %IX0.5 : BOOL;
    IN4      AT %IX0.6 : BOOL;
    IN5      AT %IX0.7 : BOOL;
    OutReady AT %QX0.0 : BOOL := FALSE;
    FeedNext AT %QX0.1 : BOOL := FALSE;
    Out      AT %QX0.2 : BOOL;
  END_VAR
  CollectInput(TICK:=TICK, IN1:=IN1, IN2:=IN2, IN3:=IN3, IN4:=IN4, IN5:=IN5);
  Ready := CollectInput.Finished;
  FeedNext := 1;
  IF Ready THEN
    Out := ((NOT Data[26]) AND (((NOT Data[23]) XOR (NOT (NOT (((((((NOT Data[29]) OR (NOT Data[21])) XOR ((((TRUE XOR Data[46]) XOR Data[14]) XOR (NOT Data[7])) XOR (NOT Data[19]))) XOR (NOT Data[12])) AND ((NOT (NOT Data[9])) OR Data[10])) OR (NOT (Data[29] AND Data[6]))) AND (((Data[34] XOR Data[46]) XOR (NOT ((Data[47] OR Data[39]) AND ((Data[48] XOR Data[16]) XOR Data[35])))) OR ((((((Data[18] XOR (NOT Data[46])) XOR Data[4]) XOR (FALSE AND (NOT Data[20]))) XOR (NOT (NOT Data[26]))) XOR FALSE) XOR (Data[34] OR ((((Data[48] XOR Data[50]) XOR Data[49]) XOR (NOT Data[38])) XOR (Data[45] AND Data[13]))))))))) XOR (((((NOT ((NOT ((FALSE XOR (NOT Data[30])) XOR Data[27])) OR (((((Data[25] AND Data[4]) XOR (Data[3] OR Data[3])) XOR (Data[47] AND Data[26])) XOR (NOT (Data[25] AND Data[25]))) XOR (NOT (NOT Data[24]))))) OR (((NOT (Data[21] OR (Data[5] AND Data[39]))) AND ((((Data[3] AND Data[24]) XOR (Data[49] AND Data[44])) XOR (Data[24] AND Data[39])) OR ((Data[21] OR Data[27]) AND Data[42]))) AND (((((NOT Data[46]) AND ((Data[42] XOR Data[44]) XOR Data[38])) AND FALSE) XOR (((((Data[38] AND FALSE) XOR Data[32]) XOR (NOT Data[21])) XOR (((Data[22] XOR Data[10]) XOR Data[42]) AND (FALSE OR Data[15]))) XOR Data[12])) XOR (((Data[22] OR (Data[41] OR Data[39])) XOR ((Data[23] OR Data[41]) AND (Data[23] AND Data[21]))) XOR ((NOT Data[22]) OR ((Data[47] XOR Data[35]) XOR Data[37])))))) XOR (((NOT ((((Data[13] AND Data[38]) OR (NOT Data[21])) OR Data[42]) OR (((Data[34] AND Data[31]) OR (Data[6] AND Data[28])) OR ((Data[45] AND Data[33]) OR Data[42])))) XOR ((Data[1] XOR ((((Data[32] AND Data[43]) AND (Data[10] OR Data[49])) AND ((((Data[42] XOR Data[8]) XOR Data[40]) XOR (Data[12] OR Data[31])) XOR (Data[25] AND Data[30]))) OR Data[13])) XOR (((((FALSE AND (Data[14] AND Data[9])) XOR (NOT Data[3])) XOR (Data[39] AND (Data[11] AND Data[35]))) XOR (Data[27] OR (NOT (Data[6] OR Data[39])))) XOR (NOT (((NOT Data[37]) XOR ((Data[1] XOR Data[13]) XOR Data[25])) XOR ((Data[22] XOR FALSE) XOR Data[17])))))) XOR (Data[31] OR (((((NOT Data[11]) AND ((Data[10] XOR Data[29]) XOR Data[38])) OR ((Data[20] AND Data[29]) OR (NOT Data[22]))) XOR Data[19]) XOR ((((Data[1] OR Data[39]) OR Data[22]) XOR ((NOT Data[7]) AND (Data[26] OR Data[10]))) XOR Data[12]))))) XOR (NOT (((NOT Data[9]) XOR (((Data[38] AND (NOT Data[35])) AND (NOT (Data[32] OR Data[20]))) AND ((TRUE XOR ((Data[35] XOR (Data[33] OR Data[35])) XOR (Data[10] OR Data[17]))) XOR (Data[42] AND ((Data[28] XOR Data[5]) XOR Data[11]))))) XOR (Data[27] AND (Data[1] OR ((NOT Data[45]) AND (Data[8] AND Data[17]))))))) OR (NOT (NOT Data[22])))));
    OutReady := 1;
    CollectInput(RESET:=TRUE);
  END_IF;
END_PROGRAM

CONFIGURATION Config0
  RESOURCE Res0 ON PLC
    TASK task0(INTERVAL := T#20ms,PRIORITY := 0);
    PROGRAM instance0 WITH task0 : Boiler;
  END_RESOURCE
END_CONFIGURATION

(* ---- RND-EXPR_yards-salsa-fiche.st ---- *)
(*
This code implements a randomly grown symbolic expression:

IN21 & IN24

*)

FUNCTION_BLOCK F_CollectInput
  VAR_IN_OUT
      Data : ARRAY[1..50] OF BOOL;
  END_VAR
  VAR_INPUT
      TICK  : BOOL := 0;
      IN1   : BOOL := 0;
      IN2   : BOOL := 0;
      IN3   : BOOL := 0;
      IN4   : BOOL := 0;
      IN5   : BOOL := 0;
      RESET : BOOL := FALSE;
  END_VAR
  VAR_OUTPUT
      Finished : BOOL;
  END_VAR
  VAR
      j    : USINT := 1;
      tock : BOOL  := 0;
  END_VAR
  IF NOT RESET AND tock = NOT TICK THEN
      Data[j]   := IN1;
      Data[j+1] := IN2;
      Data[j+2] := IN3;
      Data[j+3] := IN4;
      Data[j+4] := IN5;
      j := j + 5;
      tock := TICK;
  ELSE
      j := 1;
      tock := 0;
  END_IF;
  Finished := (j > 50);
END_FUNCTION_BLOCK

PROGRAM Boiler
  VAR
    Data  : ARRAY[1..50] OF BOOL;
    Ready : BOOL;
    CollectInput : F_CollectInput;
  END_VAR
  VAR
    TICK     AT %IX1.0 : BOOL;
    IN1      AT %IX0.3 : BOOL;
    IN2      AT %IX0.4 : BOOL;
    IN3      AT %IX0.5 : BOOL;
    IN4      AT %IX0.6 : BOOL;
    IN5      AT %IX0.7 : BOOL;
    OutReady AT %QX0.0 : BOOL := FALSE;
    FeedNext AT %QX0.1 : BOOL := FALSE;
    Out      AT %QX0.2 : BOOL;
  END_VAR
  CollectInput(TICK:=TICK, IN1:=IN1, IN2:=IN2, IN3:=IN3, IN4:=IN4, IN5:=IN5);
  Ready := CollectInput.Finished;
  FeedNext := 1;
  IF Ready THEN
    Out := (Data[21] AND Data[24]);
    OutReady := 1;
    CollectInput(RESET:=TRUE);
  END_IF;
END_PROGRAM

CONFIGURATION Config0
  RESOURCE Res0 ON PLC
    TASK task0(INTERVAL := T#20ms,PRIORITY := 0);
    PROGRAM instance0 WITH task0 : Boiler;
  END_RESOURCE
END_CONFIGURATION

(* ---- RND-EXPR_yearn-sulfa-usual.st ---- *)
(*
This code implements a randomly grown symbolic expression:

((xor(xor(IN45 & (!(((xor(xor((IN12 | IN39) & (IN49 & IN44), (xor(xor(IN32, IN2), IN29)) | (!(IN23))), !(IN43))) & ((xor(xor(!(IN34), xor(xor(IN7, IN24), IN32)), IN44 & IN23)) & (!(IN26 | IN12)))) & (xor(xor(true, (!(!(IN14))) | IN32), !((IN3 | IN34) & (xor(xor(true, IN16), IN29))))))), (true & (xor(xor(!(IN12), IN38 & ((!(IN22 & IN30)) & ((IN49 & IN6) & (xor(xor(IN28, IN16), IN47))))), IN30))) | (IN20 | (!(!(xor(xor((xor(xor(IN18, IN11), IN44)) | (IN1 | IN1), !(!(IN21))), xor(xor(!(IN27), IN8 | IN35), IN10 | IN21))))))), (IN35 | (!((!(xor(xor(!(IN11), xor(xor(IN5, IN39), IN18)), IN48 | IN49))) & (xor(xor(!(IN2 & IN40), !(IN47 & IN16)), !(xor(xor(IN48, IN6), IN12))))))) & false)) & IN28) | ((!(((((xor(xor(xor(xor(xor(xor(IN26, IN40), IN46), IN25), IN34 & IN49), (!(IN22)) & (!(IN24))), IN22)) & (((IN44 | IN23) & IN20) & (!(IN14 | IN43)))) | IN43) & ((xor(xor(IN5, (xor(xor(IN37, IN49 & IN28), xor(xor(IN22, IN20), IN30))) | ((!(IN46)) | (IN7 | IN28))), (!(IN11 | IN38)) & IN28)) | (!(IN6)))) | (xor(xor(IN22, !((((xor(xor(IN22, IN46), IN13)) | (xor(xor(IN33, IN13), IN13))) & IN3) & (xor(xor((!(IN19)) & (IN23 & IN43), IN9), !(IN47 | IN16))))), xor(xor(((xor(xor(IN41 | IN8, IN31), IN20 | IN5)) & IN33) & (xor(xor(!(IN34), (IN44 | true) & (IN24 | IN13)), IN19)), !(IN24)), !(IN43)))))) & IN28)

*)

FUNCTION_BLOCK F_CollectInput
  VAR_IN_OUT
      Data : ARRAY[1..50] OF BOOL;
  END_VAR
  VAR_INPUT
      TICK  : BOOL := 0;
      IN1   : BOOL := 0;
      IN2   : BOOL := 0;
      IN3   : BOOL := 0;
      IN4   : BOOL := 0;
      IN5   : BOOL := 0;
      RESET : BOOL := FALSE;
  END_VAR
  VAR_OUTPUT
      Finished : BOOL;
  END_VAR
  VAR
      j    : USINT := 1;
      tock : BOOL  := 0;
  END_VAR
  IF NOT RESET AND tock = NOT TICK THEN
      Data[j]   := IN1;
      Data[j+1] := IN2;
      Data[j+2] := IN3;
      Data[j+3] := IN4;
      Data[j+4] := IN5;
      j := j + 5;
      tock := TICK;
  ELSE
      j := 1;
      tock := 0;
  END_IF;
  Finished := (j > 50);
END_FUNCTION_BLOCK

PROGRAM Boiler
  VAR
    Data  : ARRAY[1..50] OF BOOL;
    Ready : BOOL;
    CollectInput : F_CollectInput;
  END_VAR
  VAR
    TICK     AT %IX1.0 : BOOL;
    IN1      AT %IX0.3 : BOOL;
    IN2      AT %IX0.4 : BOOL;
    IN3      AT %IX0.5 : BOOL;
    IN4      AT %IX0.6 : BOOL;
    IN5      AT %IX0.7 : BOOL;
    OutReady AT %QX0.0 : BOOL := FALSE;
    FeedNext AT %QX0.1 : BOOL := FALSE;
    Out      AT %QX0.2 : BOOL;
  END_VAR
  CollectInput(TICK:=TICK, IN1:=IN1, IN2:=IN2, IN3:=IN3, IN4:=IN4, IN5:=IN5);
  Ready := CollectInput.Finished;
  FeedNext := 1;
  IF Ready THEN
    Out := (((((Data[45] AND (NOT ((((((Data[12] OR Data[39]) AND (Data[49] AND Data[44])) XOR (((Data[32] XOR Data[2]) XOR Data[29]) OR (NOT Data[23]))) XOR (NOT Data[43])) AND ((((NOT Data[34]) XOR ((Data[7] XOR Data[24]) XOR Data[32])) XOR (Data[44] AND Data[23])) AND (NOT (Data[26] OR Data[12])))) AND ((TRUE XOR ((NOT (NOT Data[14])) OR Data[32])) XOR (NOT ((Data[3] OR Data[34]) AND ((TRUE XOR Data[16]) XOR Data[29]))))))) XOR ((TRUE AND (((NOT Data[12]) XOR (Data[38] AND ((NOT (Data[22] AND Data[30])) AND ((Data[49] AND Data[6]) AND ((Data[28] XOR Data[16]) XOR Data[47]))))) XOR Data[30])) OR (Data[20] OR (NOT (NOT (((((Data[18] XOR Data[11]) XOR Data[44]) OR (Data[1] OR Data[1])) XOR (NOT (NOT Data[21]))) XOR (((NOT Data[27]) XOR (Data[8] OR Data[35])) XOR (Data[10] OR Data[21])))))))) XOR ((Data[35] OR (NOT ((NOT (((NOT Data[11]) XOR ((Data[5] XOR Data[39]) XOR Data[18])) XOR (Data[48] OR Data[49]))) AND (((NOT (Data[2] AND Data[40])) XOR (NOT (Data[47] AND Data[16]))) XOR (NOT ((Data[48] XOR Data[6]) XOR Data[12])))))) AND FALSE)) AND Data[28]) OR ((NOT ((((((((((Data[26] XOR Data[40]) XOR Data[46]) XOR Data[25]) XOR (Data[34] AND Data[49])) XOR ((NOT Data[22]) AND (NOT Data[24]))) XOR Data[22]) AND (((Data[44] OR Data[23]) AND Data[20]) AND (NOT (Data[14] OR Data[43])))) OR Data[43]) AND (((Data[5] XOR (((Data[37] XOR (Data[49] AND Data[28])) XOR ((Data[22] XOR Data[20]) XOR Data[30])) OR ((NOT Data[46]) OR (Data[7] OR Data[28])))) XOR ((NOT (Data[11] OR Data[38])) AND Data[28])) OR (NOT Data[6]))) OR ((Data[22] XOR (NOT (((((Data[22] XOR Data[46]) XOR Data[13]) OR ((Data[33] XOR Data[13]) XOR Data[13])) AND Data[3]) AND ((((NOT Data[19]) AND (Data[23] AND Data[43])) XOR Data[9]) XOR (NOT (Data[47] OR Data[16])))))) XOR (((((((Data[41] OR Data[8]) XOR Data[31]) XOR (Data[20] OR Data[5])) AND Data[33]) AND (((NOT Data[34]) XOR ((Data[44] OR TRUE) AND (Data[24] OR Data[13]))) XOR Data[19])) XOR (NOT Data[24])) XOR (NOT Data[43]))))) AND Data[28]));
    OutReady := 1;
    CollectInput(RESET:=TRUE);
  END_IF;
END_PROGRAM

CONFIGURATION Config0
  RESOURCE Res0 ON PLC
    TASK task0(INTERVAL := T#20ms,PRIORITY := 0);
    PROGRAM instance0 WITH task0 : Boiler;
  END_RESOURCE
END_CONFIGURATION

(* ---- RND-EXPR_astro-cried-peers.st ---- *)
(*
This code implements a randomly grown symbolic expression:

xor(xor(xor(xor(xor(xor(xor(xor((!(!(!(xor(xor(!(IN34), !(IN44)), xor(xor(IN30, IN41), IN27)))))) & (!(((IN27 & (IN10 | IN5)) | (xor(xor(false, !(IN14)), IN38 | IN43))) | ((xor(xor(xor(xor(IN1, IN34), IN14), IN29), xor(xor(IN39, IN14), IN28))) | (!(IN23))))), ((!(!((xor(xor(IN31, IN11), IN7)) | IN39))) & (!((!(IN39 | IN35)) | IN10))) & (!((IN6 | (!(!(IN31)))) | ((!(!(IN13))) & ((xor(xor(IN14, IN50), IN11)) | (xor(xor(IN21, IN31), IN33))))))), xor(xor(IN8, IN3), xor(xor(((xor(xor(IN39, xor(xor(IN31, IN28), IN34)), IN49 | IN28)) | ((IN16 | IN6) | (xor(xor(IN35, IN37), false)))) | ((xor(xor(!(IN37), xor(xor(IN27, IN42), IN3)), IN2 | IN4)) | (!(!(IN29)))), (xor(xor(!(!(IN14)), (!(IN29)) & (IN30 & IN40)), IN11)) & (IN33 | IN43)), xor(xor(xor(xor(!(IN35), !(!(IN6))), !(IN26)), xor(xor(xor(xor(!(IN44), IN24 | IN17), IN17 & IN49), !(IN8 | IN47)), !(IN31 & IN26))), xor(xor(IN44 & (!(IN27)), !(IN2 & IN27)), (!(IN23)) | IN21))))), xor(xor((!(IN1)) & (!(IN44 | IN45)), xor(xor((!((xor(xor(IN43, !(IN49)), IN2 | IN21)) | (xor(xor(IN31 & IN46, IN42 | IN4), !(IN18))))) | (xor(xor((IN8 | (!(IN33))) & IN16, IN24 & IN2), ((IN31 | IN9) & true) & (xor(xor(IN22 & IN44, IN19 & IN37), IN9 & IN6)))), (!(IN11 & (!(!(IN28))))) & (!(!(!(IN49))))), (xor(xor(((!(IN15)) & IN13) | (xor(xor(!(IN26), !(IN48)), true & IN29)), xor(xor((IN11 | IN31) | (!(IN11)), (IN20 | IN35) | (IN30 | IN49)), xor(xor(xor(xor(IN27, IN43), IN9), IN6 | IN35), IN17 & IN7))), !(xor(xor(!(IN37), xor(xor(IN39, false), false)), xor(xor(IN11, IN45), IN44))))) & (IN10 | ((xor(xor(IN1 | IN5, !(IN36)), !(IN21))) & (xor(xor(!(IN27), IN16), xor(xor(IN7, false), IN48))))))), IN3 & (xor(xor((IN4 | IN30) | (!(IN35 & (false & IN19))), xor(xor(((xor(xor(IN48, IN15), IN9)) & (IN47 | IN26)) | IN27, xor(xor(xor(xor(IN41 & IN10, xor(xor(IN39, true), IN9)), xor(xor(IN12, IN47), IN32)), xor(xor(IN5 | IN18, IN4 | IN3), IN12 | IN35)), !(IN49))), !((IN8 & IN4) | (xor(xor(IN5, IN12), IN32))))), !(IN45 | IN22))))), xor(xor(!(((!((IN10 | IN4) & (!(IN43)))) | IN32) | ((xor(xor(xor(xor(false, IN4 & IN41), IN20 | IN32), IN33 | (xor(xor(IN37, false), IN21))), xor(xor(IN29 & IN4, xor(xor(IN12, IN18), IN39)), IN7 | IN31))) | (!(xor(xor(IN22 & IN16, xor(xor(IN17, IN22), IN33)), !(IN29)))))), IN13), !(xor(xor((((IN33 & IN40) & (xor(xor(IN24, IN45), IN25))) & ((IN25 | IN42) | (IN17 & IN9))) & (IN48 | (!(xor(xor(IN41, IN11), IN1)))), !(IN41)), ((xor(xor(xor(xor(IN13, IN27), IN12), IN35 | IN18), xor(xor(IN20, IN15), IN29))) | (!(!(IN7)))) | ((true | (IN17 | IN47)) | (!(xor(xor(IN29, IN7), IN47)))))))), IN12), xor(xor(IN26 & (xor(xor(xor(xor(IN19, xor(xor(xor(xor(xor(xor(IN24, IN50 & IN2), !(IN42)), xor(xor(IN40 & IN5, IN10 | IN14), IN34 | IN14)), IN44), xor(xor((xor(xor(IN7, IN45), IN46)) & IN30, (!(IN47)) | (IN39 & true)), xor(xor(IN9 | IN50, true), IN26))), (xor(xor(!(IN12), IN6 & IN3), xor(xor(IN47, IN15), IN30))) & (xor(xor(xor(xor(IN18, IN35), IN49), IN32), IN46 | IN32)))), IN4), IN43 | ((!(!(!(IN12)))) | (((IN38 & IN10) & (!(IN33))) & false))), xor(xor(!((xor(xor(IN47 | IN27, !(IN21)), IN35 | IN6)) | ((!(IN45)) | (!(IN1)))), ((xor(xor(xor(xor(IN33, IN30), IN3), IN48), IN10)) | ((!(IN34)) & IN5)) | (!(IN42))), IN5))), xor(xor(IN21, xor(xor(xor(xor((((xor(xor(IN2, IN5), IN39)) | (IN16 & IN23)) | ((IN32 | IN47) | (IN16 | IN50))) & ((!(!(IN18))) | (true | (xor(xor(IN9, IN46), IN13)))), xor(xor(IN28, (xor(xor(IN9, xor(xor(IN41, IN31), IN22)), IN36)) | (xor(xor(!(IN20), IN2 | IN3), xor(xor(IN36, IN47), IN46)))), ((IN26 & IN33) | (IN39 & IN22)) | (!(!(IN9))))), (!(!(IN26 | IN31))) | (xor(xor(IN27, (xor(xor(IN22, IN8), IN5)) | (IN12 & IN15)), !(IN21 | IN8)))), xor(xor(!(IN26 | IN21), (!(!(IN19))) & ((!(IN35 & IN21)) & (xor(xor(false, IN1 & IN44), IN19 | IN14)))), xor(xor((xor(xor(IN8 | IN22, IN27 | IN12), !(IN27))) | IN32, !((!(IN11)) & (IN10 | IN44))), IN24))), ((xor(xor(IN33, xor(xor(xor(xor(IN2, IN43), IN21), IN31 | IN37), IN11 | IN18)), xor(xor(IN18, IN41), IN44 | IN3))) | IN30) & (!(xor(xor((!(IN45)) & (IN1 & IN37), xor(xor(IN17 & IN14, IN28 | IN49), !(IN26))), (xor(xor(IN42, IN5), IN35)) & (IN27 | IN3)))))), (IN3 | ((xor(xor(IN23, IN27), (xor(xor(IN15, IN4), IN15)) & (xor(xor(IN12, IN14), IN38)))) | (xor(xor(!(IN31), (!(IN12)) & IN33), IN40)))) & ((!(xor(xor(IN14 | (IN49 & IN32), true | (!(IN24))), xor(xor(!(IN6), IN44 & IN7), IN13)))) & (((!(IN23 & IN46)) | false) & ((xor(xor(IN35 & IN25, IN31 | IN15), !(IN30))) | ((IN28 & IN38) & (IN27 & false))))))), (((xor(xor(!(xor(xor(IN25 & IN45, !(IN18)), xor(xor(IN27, IN41), IN15))), xor(xor(!(IN33), (IN46 | IN50) & (IN15 & IN37)), IN45)), (IN39 & (!(IN16))) | ((!(IN29)) | (!(IN47))))) & (xor(xor(IN42, (xor(xor(!(IN42), xor(xor(IN23, IN26), IN5)), IN24 & IN28)) | ((IN49 | IN8) | (xor(xor(IN21, IN15), IN30)))), false))) | ((xor(xor((IN24 | (xor(xor(IN48, IN23), IN28))) | (IN32 | IN25), ((IN17 | IN16) | (!(IN6))) | (!(IN13 & IN11))), (xor(xor(IN46 | IN19, IN26), IN42 & IN27)) & (IN15 & (IN21 & IN46)))) & (!(xor(xor(!(xor(xor(IN34, IN6), IN31)), !(IN40 | IN5)), xor(xor(IN28 | IN9, xor(xor(IN21, IN27), IN36)), IN10 | IN6)))))) | (!(IN41)))), IN29), xor(xor((xor(xor(IN11, (((((IN18 | IN13) | (xor(xor(IN21, IN11), IN16))) | (!(IN3 & IN2))) & (xor(true, !(IN4 & IN7)))) & IN26) & (xor(xor(xor(xor(xor(xor((IN8 & IN42) | (IN35 | IN7), !(IN43 | IN43)), (IN38 & IN30) & (IN6 & IN24)), (!(IN30)) & (!(IN8 & IN26))), IN46), xor(xor(xor(xor(IN18 | (xor(xor(IN18, IN8), IN48)), !(IN32)), (!(IN13)) & IN1), !(xor(xor(IN36 & IN39, IN31), IN1 | IN43))), IN28)), (xor(xor(IN14 & (IN28 & IN41), (IN26 & IN15) & (IN15 | IN21)), (IN29 | IN9) | (IN30 | IN38))) & (!((IN5 & IN24) | (!(IN46))))))), IN43)) & (((((!(xor(xor(!(IN17), IN18 | IN16), xor(xor(IN34, IN1), IN31)))) & (IN44 | IN11)) | (IN19 & (IN13 & IN23))) | (!(xor(xor(!(IN25), xor(xor((IN7 | IN34) | (IN36 | IN30), (IN17 | IN2) & (!(IN23))), IN46)), xor(xor(xor(xor(IN27, xor(xor(IN15, IN32), IN23)), IN29), !(!(IN49))), IN1))))) | false), ((IN22 & ((!(IN13)) & ((!((IN33 & false) & (IN7 | IN28))) | IN41))) & (IN32 & (((IN3 | (!(IN27 & IN13))) | (!((IN26 & IN3) & (xor(xor(IN41, IN35), IN44))))) | IN18))) & ((xor(xor((xor(xor(!((xor(xor(IN15, IN34), true)) | (IN17 | IN36)), IN26 | (!(xor(xor(IN50, IN5), IN45)))), !(xor(xor(IN44 & IN27, xor(xor(IN18, IN42), IN27)), IN24 | IN23)))) | (!(xor(xor(!(!(IN47)), xor(xor(xor(xor(IN23, IN37), IN6), IN41 & IN29), !(IN48))), (IN36 | IN20) | (!(IN32))))), (xor(xor((xor(xor(IN7 & IN37, IN29 | IN23), IN18 & IN40)) & ((IN34 & IN26) & (IN28 | IN49)), xor(xor(xor(xor(IN20, IN34 & IN28), IN6 | IN46), (xor(xor(IN8, IN7), IN22)) | (IN1 | IN16)), (xor(xor(IN1, IN36), IN2)) | (!(IN47)))), !((xor(xor(IN27, IN18), IN37)) | (!(IN40))))) | IN31), (!(IN30 | ((IN47 | IN18) & IN29))) & (xor(xor((!(!(IN17))) | (!(IN38)), IN11), ((xor(xor(IN34, IN25), IN37)) & (true & IN36)) & ((!(IN45)) | (IN14 & IN37)))))) & ((xor(xor(IN12, !(IN47)), !(IN16 & (xor(xor(!(IN32), xor(xor(IN37, IN35), IN28)), IN38 | IN13))))) | (!(IN15 | IN39))))), (((!(!(!(IN3)))) & (((!((IN13 | IN47) | (xor(xor(IN11, IN45), IN37)))) & (IN21 & IN14)) & ((((IN12 | IN17) & (xor(xor(IN12, IN13), IN4))) | (!(!(IN37)))) & IN26))) & (xor(xor(IN48, xor(xor(IN41, xor(xor(IN22, ((IN35 & IN36) | false) & (!(IN10 | IN37))), (!(IN9)) | ((xor(xor(IN12, IN21), IN31)) & (!(IN12))))), !(IN22))), xor(xor(xor(xor(IN37 | ((!(IN47)) & IN12), xor(xor((IN15 & IN44) | (!(IN12)), !(IN28 | IN39)), IN36)), !(IN26 & false)), !(!(!(!(IN40))))), IN20)))) & ((((((!(IN5 & IN21)) | (!(xor(xor(IN28, IN45), IN33)))) & (!(xor(xor(xor(xor(IN18, IN50), IN8), !(IN15)), IN10 | IN47)))) & (((xor(xor(IN19 | IN50, IN43), xor(xor(IN50, IN17), IN36))) | IN25) & (!(xor(xor(xor(xor(IN12, IN28), IN25), IN8), IN48 & IN2))))) & (!((!(!(!(IN50)))) | IN11))) | (!((!(((true | IN28) | (false | IN48)) | ((!(IN11)) | (IN38 & IN41)))) & ((IN15 & (xor(xor(IN31, !(IN37)), IN16 | IN8))) | (xor(xor(IN46, !(!(IN19))), (IN14 | IN8) | (IN21 | IN14)))))))))

*)

FUNCTION_BLOCK F_CollectInput
  VAR_IN_OUT
      Data : ARRAY[1..50] OF BOOL;
  END_VAR
  VAR_INPUT
      TICK  : BOOL := 0;
      IN1   : BOOL := 0;
      IN2   : BOOL := 0;
      IN3   : BOOL := 0;
      IN4   : BOOL := 0;
      IN5   : BOOL := 0;
      RESET : BOOL := FALSE;
  END_VAR
  VAR_OUTPUT
      Finished : BOOL;
  END_VAR
  VAR
      j    : USINT := 1;
      tock : BOOL  := 0;
  END_VAR
  IF NOT RESET AND tock = NOT TICK THEN
      Data[j]   := IN1;
      Data[j+1] := IN2;
      Data[j+2] := IN3;
      Data[j+3] := IN4;
      Data[j+4] := IN5;
      j := j + 5;
      tock := TICK;
  ELSE
      j := 1;
      tock := 0;
  END_IF;
  Finished := (j > 50);
END_FUNCTION_BLOCK

PROGRAM Boiler
  VAR
    Data  : ARRAY[1..50] OF BOOL;
    Ready : BOOL;
    CollectInput : F_CollectInput;
  END_VAR
  VAR
    TICK     AT %IX1.0 : BOOL;
    IN1      AT %IX0.3 : BOOL;
    IN2      AT %IX0.4 : BOOL;
    IN3      AT %IX0.5 : BOOL;
    IN4      AT %IX0.6 : BOOL;
    IN5      AT %IX0.7 : BOOL;
    OutReady AT %QX0.0 : BOOL := FALSE;
    FeedNext AT %QX0.1 : BOOL := FALSE;
    Out      AT %QX0.2 : BOOL;
  END_VAR
  CollectInput(TICK:=TICK, IN1:=IN1, IN2:=IN2, IN3:=IN3, IN4:=IN4, IN5:=IN5);
  Ready := CollectInput.Finished;
  FeedNext := 1;
  IF Ready THEN
    Out := ((((((((((NOT (NOT (NOT (((NOT Data[34]) XOR (NOT Data[44])) XOR ((Data[30] XOR Data[41]) XOR Data[27]))))) AND (NOT (((Data[27] AND (Data[10] OR Data[5])) OR ((FALSE XOR (NOT Data[14])) XOR (Data[38] OR Data[43]))) OR (((((Data[1] XOR Data[34]) XOR Data[14]) XOR Data[29]) XOR ((Data[39] XOR Data[14]) XOR Data[28])) OR (NOT Data[23]))))) XOR (((NOT (NOT (((Data[31] XOR Data[11]) XOR Data[7]) OR Data[39]))) AND (NOT ((NOT (Data[39] OR Data[35])) OR Data[10]))) AND (NOT ((Data[6] OR (NOT (NOT Data[31]))) OR ((NOT (NOT Data[13])) AND (((Data[14] XOR Data[50]) XOR Data[11]) OR ((Data[21] XOR Data[31]) XOR Data[33]))))))) XOR ((Data[8] XOR Data[3]) XOR ((((((Data[39] XOR ((Data[31] XOR Data[28]) XOR Data[34])) XOR (Data[49] OR Data[28])) OR ((Data[16] OR Data[6]) OR ((Data[35] XOR Data[37]) XOR FALSE))) OR ((((NOT Data[37]) XOR ((Data[27] XOR Data[42]) XOR Data[3])) XOR (Data[2] OR Data[4])) OR (NOT (NOT Data[29])))) XOR ((((NOT (NOT Data[14])) XOR ((NOT Data[29]) AND (Data[30] AND Data[40]))) XOR Data[11]) AND (Data[33] OR Data[43]))) XOR (((((NOT Data[35]) XOR (NOT (NOT Data[6]))) XOR (NOT Data[26])) XOR (((((NOT Data[44]) XOR (Data[24] OR Data[17])) XOR (Data[17] AND Data[49])) XOR (NOT (Data[8] OR Data[47]))) XOR (NOT (Data[31] AND Data[26])))) XOR (((Data[44] AND (NOT Data[27])) XOR (NOT (Data[2] AND Data[27]))) XOR ((NOT Data[23]) OR Data[21])))))) XOR ((((NOT Data[1]) AND (NOT (Data[44] OR Data[45]))) XOR ((((NOT (((Data[43] XOR (NOT Data[49])) XOR (Data[2] OR Data[21])) OR (((Data[31] AND Data[46]) XOR (Data[42] OR Data[4])) XOR (NOT Data[18])))) OR ((((Data[8] OR (NOT Data[33])) AND Data[16]) XOR (Data[24] AND Data[2])) XOR (((Data[31] OR Data[9]) AND TRUE) AND (((Data[22] AND Data[44]) XOR (Data[19] AND Data[37])) XOR (Data[9] AND Data[6]))))) XOR ((NOT (Data[11] AND (NOT (NOT Data[28])))) AND (NOT (NOT (NOT Data[49]))))) XOR ((((((NOT Data[15]) AND Data[13]) OR (((NOT Data[26]) XOR (NOT Data[48])) XOR (TRUE AND Data[29]))) XOR ((((Data[11] OR Data[31]) OR (NOT Data[11])) XOR ((Data[20] OR Data[35]) OR (Data[30] OR Data[49]))) XOR ((((Data[27] XOR Data[43]) XOR Data[9]) XOR (Data[6] OR Data[35])) XOR (Data[17] AND Data[7])))) XOR (NOT (((NOT Data[37]) XOR ((Data[39] XOR FALSE) XOR FALSE)) XOR ((Data[11] XOR Data[45]) XOR Data[44])))) AND (Data[10] OR ((((Data[1] OR Data[5]) XOR (NOT Data[36])) XOR (NOT Data[21])) AND (((NOT Data[27]) XOR Data[16]) XOR ((Data[7] XOR FALSE) XOR Data[48]))))))) XOR (Data[3] AND ((((Data[4] OR Data[30]) OR (NOT (Data[35] AND (FALSE AND Data[19])))) XOR ((((((Data[48] XOR Data[15]) XOR Data[9]) AND (Data[47] OR Data[26])) OR Data[27]) XOR (((((Data[41] AND Data[10]) XOR ((Data[39] XOR TRUE) XOR Data[9])) XOR ((Data[12] XOR Data[47]) XOR Data[32])) XOR (((Data[5] OR Data[18]) XOR (Data[4] OR Data[3])) XOR (Data[12] OR Data[35]))) XOR (NOT Data[49]))) XOR (NOT ((Data[8] AND Data[4]) OR ((Data[5] XOR Data[12]) XOR Data[32]))))) XOR (NOT (Data[45] OR Data[22])))))) XOR (((NOT (((NOT ((Data[10] OR Data[4]) AND (NOT Data[43]))) OR Data[32]) OR (((((FALSE XOR (Data[4] AND Data[41])) XOR (Data[20] OR Data[32])) XOR (Data[33] OR ((Data[37] XOR FALSE) XOR Data[21]))) XOR (((Data[29] AND Data[4]) XOR ((Data[12] XOR Data[18]) XOR Data[39])) XOR (Data[7] OR Data[31]))) OR (NOT (((Data[22] AND Data[16]) XOR ((Data[17] XOR Data[22]) XOR Data[33])) XOR (NOT Data[29])))))) XOR Data[13]) XOR (NOT ((((((Data[33] AND Data[40]) AND ((Data[24] XOR Data[45]) XOR Data[25])) AND ((Data[25] OR Data[42]) OR (Data[17] AND Data[9]))) AND (Data[48] OR (NOT ((Data[41] XOR Data[11]) XOR Data[1])))) XOR (NOT Data[41])) XOR ((((((Data[13] XOR Data[27]) XOR Data[12]) XOR (Data[35] OR Data[18])) XOR ((Data[20] XOR Data[15]) XOR Data[29])) OR (NOT (NOT Data[7]))) OR ((TRUE OR (Data[17] OR Data[47])) OR (NOT ((Data[29] XOR Data[7]) XOR Data[47])))))))) XOR Data[12]) XOR (((Data[26] AND ((((Data[19] XOR ((((((Data[24] XOR (Data[50] AND Data[2])) XOR (NOT Data[42])) XOR (((Data[40] AND Data[5]) XOR (Data[10] OR Data[14])) XOR (Data[34] OR Data[14]))) XOR Data[44]) XOR (((((Data[7] XOR Data[45]) XOR Data[46]) AND Data[30]) XOR ((NOT Data[47]) OR (Data[39] AND TRUE))) XOR (((Data[9] OR Data[50]) XOR TRUE) XOR Data[26]))) XOR ((((NOT Data[12]) XOR (Data[6] AND Data[3])) XOR ((Data[47] XOR Data[15]) XOR Data[30])) AND ((((Data[18] XOR Data[35]) XOR Data[49]) XOR Data[32]) XOR (Data[46] OR Data[32]))))) XOR Data[4]) XOR (Data[43] OR ((NOT (NOT (NOT Data[12]))) OR (((Data[38] AND Data[10]) AND (NOT Data[33])) AND FALSE)))) XOR (((NOT ((((Data[47] OR Data[27]) XOR (NOT Data[21])) XOR (Data[35] OR Data[6])) OR ((NOT Data[45]) OR (NOT Data[1])))) XOR ((((((Data[33] XOR Data[30]) XOR Data[3]) XOR Data[48]) XOR Data[10]) OR ((NOT Data[34]) AND Data[5])) OR (NOT Data[42]))) XOR Data[5]))) XOR ((Data[21] XOR (((((((((Data[2] XOR Data[5]) XOR Data[39]) OR (Data[16] AND Data[23])) OR ((Data[32] OR Data[47]) OR (Data[16] OR Data[50]))) AND ((NOT (NOT Data[18])) OR (TRUE OR ((Data[9] XOR Data[46]) XOR Data[13])))) XOR ((Data[28] XOR (((Data[9] XOR ((Data[41] XOR Data[31]) XOR Data[22])) XOR Data[36]) OR (((NOT Data[20]) XOR (Data[2] OR Data[3])) XOR ((Data[36] XOR Data[47]) XOR Data[46])))) XOR (((Data[26] AND Data[33]) OR (Data[39] AND Data[22])) OR (NOT (NOT Data[9]))))) XOR ((NOT (NOT (Data[26] OR Data[31]))) OR ((Data[27] XOR (((Data[22] XOR Data[8]) XOR Data[5]) OR (Data[12] AND Data[15]))) XOR (NOT (Data[21] OR Data[8]))))) XOR (((NOT (Data[26] OR Data[21])) XOR ((NOT (NOT Data[19])) AND ((NOT (Data[35] AND Data[21])) AND ((FALSE XOR (Data[1] AND Data[44])) XOR (Data[19] OR Data[14]))))) XOR ((((((Data[8] OR Data[22]) XOR (Data[27] OR Data[12])) XOR (NOT Data[27])) OR Data[32]) XOR (NOT ((NOT Data[11]) AND (Data[10] OR Data[44])))) XOR Data[24]))) XOR ((((Data[33] XOR ((((Data[2] XOR Data[43]) XOR Data[21]) XOR (Data[31] OR Data[37])) XOR (Data[11] OR Data[18]))) XOR ((Data[18] XOR Data[41]) XOR (Data[44] OR Data[3]))) OR Data[30]) AND (NOT ((((NOT Data[45]) AND (Data[1] AND Data[37])) XOR (((Data[17] AND Data[14]) XOR (Data[28] OR Data[49])) XOR (NOT Data[26]))) XOR (((Data[42] XOR Data[5]) XOR Data[35]) AND (Data[27] OR Data[3]))))))) XOR ((Data[3] OR (((Data[23] XOR Data[27]) XOR (((Data[15] XOR Data[4]) XOR Data[15]) AND ((Data[12] XOR Data[14]) XOR Data[38]))) OR (((NOT Data[31]) XOR ((NOT Data[12]) AND Data[33])) XOR Data[40]))) AND ((NOT (((Data[14] OR (Data[49] AND Data[32])) XOR (TRUE OR (NOT Data[24]))) XOR (((NOT Data[6]) XOR (Data[44] AND Data[7])) XOR Data[13]))) AND (((NOT (Data[23] AND Data[46])) OR FALSE) AND ((((Data[35] AND Data[25]) XOR (Data[31] OR Data[15])) XOR (NOT Data[30])) OR ((Data[28] AND Data[38]) AND (Data[27] AND FALSE)))))))) XOR ((((((NOT (((Data[25] AND Data[45]) XOR (NOT Data[18])) XOR ((Data[27] XOR Data[41]) XOR Data[15]))) XOR (((NOT Data[33]) XOR ((Data[46] OR Data[50]) AND (Data[15] AND Data[37]))) XOR Data[45])) XOR ((Data[39] AND (NOT Data[16])) OR ((NOT Data[29]) OR (NOT Data[47])))) AND ((Data[42] XOR ((((NOT Data[42]) XOR ((Data[23] XOR Data[26]) XOR Data[5])) XOR (Data[24] AND Data[28])) OR ((Data[49] OR Data[8]) OR ((Data[21] XOR Data[15]) XOR Data[30])))) XOR FALSE)) OR (((((Data[24] OR ((Data[48] XOR Data[23]) XOR Data[28])) OR (Data[32] OR Data[25])) XOR (((Data[17] OR Data[16]) OR (NOT Data[6])) OR (NOT (Data[13] AND Data[11])))) XOR ((((Data[46] OR Data[19]) XOR Data[26]) XOR (Data[42] AND Data[27])) AND (Data[15] AND (Data[21] AND Data[46])))) AND (NOT (((NOT ((Data[34] XOR Data[6]) XOR Data[31])) XOR (NOT (Data[40] OR Data[5]))) XOR (((Data[28] OR Data[9]) XOR ((Data[21] XOR Data[27]) XOR Data[36])) XOR (Data[10] OR Data[6])))))) OR (NOT Data[41])))) XOR Data[29]) XOR (((((Data[11] XOR ((((((Data[18] OR Data[13]) OR ((Data[21] XOR Data[11]) XOR Data[16])) OR (NOT (Data[3] AND Data[2]))) AND (TRUE XOR (NOT (Data[4] AND Data[7])))) AND Data[26]) AND ((((((((Data[8] AND Data[42]) OR (Data[35] OR Data[7])) XOR (NOT (Data[43] OR Data[43]))) XOR ((Data[38] AND Data[30]) AND (Data[6] AND Data[24]))) XOR ((NOT Data[30]) AND (NOT (Data[8] AND Data[26])))) XOR Data[46]) XOR (((((Data[18] OR ((Data[18] XOR Data[8]) XOR Data[48])) XOR (NOT Data[32])) XOR ((NOT Data[13]) AND Data[1])) XOR (NOT (((Data[36] AND Data[39]) XOR Data[31]) XOR (Data[1] OR Data[43])))) XOR Data[28])) XOR ((((Data[14] AND (Data[28] AND Data[41])) XOR ((Data[26] AND Data[15]) AND (Data[15] OR Data[21]))) XOR ((Data[29] OR Data[9]) OR (Data[30] OR Data[38]))) AND (NOT ((Data[5] AND Data[24]) OR (NOT Data[46]))))))) XOR Data[43]) AND (((((NOT (((NOT Data[17]) XOR (Data[18] OR Data[16])) XOR ((Data[34] XOR Data[1]) XOR Data[31]))) AND (Data[44] OR Data[11])) OR (Data[19] AND (Data[13] AND Data[23]))) OR (NOT (((NOT Data[25]) XOR ((((Data[7] OR Data[34]) OR (Data[36] OR Data[30])) XOR ((Data[17] OR Data[2]) AND (NOT Data[23]))) XOR Data[46])) XOR ((((Data[27] XOR ((Data[15] XOR Data[32]) XOR Data[23])) XOR Data[29]) XOR (NOT (NOT Data[49]))) XOR Data[1])))) OR FALSE)) XOR (((Data[22] AND ((NOT Data[13]) AND ((NOT ((Data[33] AND FALSE) AND (Data[7] OR Data[28]))) OR Data[41]))) AND (Data[32] AND (((Data[3] OR (NOT (Data[27] AND Data[13]))) OR (NOT ((Data[26] AND Data[3]) AND ((Data[41] XOR Data[35]) XOR Data[44])))) OR Data[18]))) AND (((((((NOT (((Data[15] XOR Data[34]) XOR TRUE) OR (Data[17] OR Data[36]))) XOR (Data[26] OR (NOT ((Data[50] XOR Data[5]) XOR Data[45])))) XOR (NOT (((Data[44] AND Data[27]) XOR ((Data[18] XOR Data[42]) XOR Data[27])) XOR (Data[24] OR Data[23])))) OR (NOT (((NOT (NOT Data[47])) XOR ((((Data[23] XOR Data[37]) XOR Data[6]) XOR (Data[41] AND Data[29])) XOR (NOT Data[48]))) XOR ((Data[36] OR Data[20]) OR (NOT Data[32]))))) XOR (((((((Data[7] AND Data[37]) XOR (Data[29] OR Data[23])) XOR (Data[18] AND Data[40])) AND ((Data[34] AND Data[26]) AND (Data[28] OR Data[49]))) XOR ((((Data[20] XOR (Data[34] AND Data[28])) XOR (Data[6] OR Data[46])) XOR (((Data[8] XOR Data[7]) XOR Data[22]) OR (Data[1] OR Data[16]))) XOR (((Data[1] XOR Data[36]) XOR Data[2]) OR (NOT Data[47])))) XOR (NOT (((Data[27] XOR Data[18]) XOR Data[37]) OR (NOT Data[40])))) OR Data[31])) XOR ((NOT (Data[30] OR ((Data[47] OR Data[18]) AND Data[29]))) AND ((((NOT (NOT Data[17])) OR (NOT Data[38])) XOR Data[11]) XOR ((((Data[34] XOR Data[25]) XOR Data[37]) AND (TRUE AND Data[36])) AND ((NOT Data[45]) OR (Data[14] AND Data[37])))))) AND (((Data[12] XOR (NOT Data[47])) XOR (NOT (Data[16] AND (((NOT Data[32]) XOR ((Data[37] XOR Data[35]) XOR Data[28])) XOR (Data[38] OR Data[13]))))) OR (NOT (Data[15] OR Data[39])))))) XOR ((((NOT (NOT (NOT Data[3]))) AND (((NOT ((Data[13] OR Data[47]) OR ((Data[11] XOR Data[45]) XOR Data[37]))) AND (Data[21] AND Data[14])) AND ((((Data[12] OR Data[17]) AND ((Data[12] XOR Data[13]) XOR Data[4])) OR (NOT (NOT Data[37]))) AND Data[26]))) AND ((Data[48] XOR ((Data[41] XOR ((Data[22] XOR (((Data[35] AND Data[36]) OR FALSE) AND (NOT (Data[10] OR Data[37])))) XOR ((NOT Data[9]) OR (((Data[12] XOR Data[21]) XOR Data[31]) AND (NOT Data[12]))))) XOR (NOT Data[22]))) XOR (((((Data[37] OR ((NOT Data[47]) AND Data[12])) XOR ((((Data[15] AND Data[44]) OR (NOT Data[12])) XOR (NOT (Data[28] OR Data[39]))) XOR Data[36])) XOR (NOT (Data[26] AND FALSE))) XOR (NOT (NOT (NOT (NOT Data[40]))))) XOR Data[20]))) AND ((((((NOT (Data[5] AND Data[21])) OR (NOT ((Data[28] XOR Data[45]) XOR Data[33]))) AND (NOT ((((Data[18] XOR Data[50]) XOR Data[8]) XOR (NOT Data[15])) XOR (Data[10] OR Data[47])))) AND (((((Data[19] OR Data[50]) XOR Data[43]) XOR ((Data[50] XOR Data[17]) XOR Data[36])) OR Data[25]) AND (NOT ((((Data[12] XOR Data[28]) XOR Data[25]) XOR Data[8]) XOR (Data[48] AND Data[2]))))) AND (NOT ((NOT (NOT (NOT Data[50]))) OR Data[11]))) OR (NOT ((NOT (((TRUE OR Data[28]) OR (FALSE OR Data[48])) OR ((NOT Data[11]) OR (Data[38] AND Data[41])))) AND ((Data[15] AND ((Data[31] XOR (NOT Data[37])) XOR (Data[16] OR Data[8]))) OR ((Data[46] XOR (NOT (NOT Data[19]))) XOR ((Data[14] OR Data[8]) OR (Data[21] OR Data[14]))))))))));
    OutReady := 1;
    CollectInput(RESET:=TRUE);
  END_IF;
END_PROGRAM

CONFIGURATION Config0
  RESOURCE Res0 ON PLC
    TASK task0(INTERVAL := T#20ms,PRIORITY := 0);
    PROGRAM instance0 WITH task0 : Boiler;
  END_RESOURCE
END_CONFIGURATION

(* ---- RND-EXPR_built-lasts-soaps.st ---- *)
(*
This code implements a randomly grown symbolic expression:

(xor(xor(!(IN49), IN20), !(!((!(!(IN20))) | ((!(((IN1 | IN21) & (xor(xor(IN13, IN2), IN39))) & (!(IN34 | IN7)))) & (!(!(xor(xor(IN4 & IN42, xor(xor(IN12, IN33), IN1)), !(IN24)))))))))) | (xor(xor(xor(xor(xor(xor(((xor(xor(!(!(IN2 & IN8)), ((IN41 & IN1) & (IN10 | IN13)) & IN47), !((xor(xor(IN42, IN37), IN36)) & IN20))) & true) | IN48, IN37), (!((!((xor(xor(IN26, IN18), IN46)) | (IN49 & IN34))) | (((xor(xor(IN3, IN49), IN16)) | (!(IN33))) | IN21))) & (xor(xor((!(xor(xor(false | IN24, !(IN1)), xor(xor(IN46, IN37), IN21)))) & (!(IN49)), IN13), !(xor(xor((IN41 | IN32) | IN21, (xor(xor(IN18, IN1), IN35)) | (xor(xor(IN21, IN7), IN35))), (!(IN41)) & (IN27 & IN20)))))), (((((IN50 & (xor(xor(IN19, IN26), IN19))) & ((!(IN47)) & (xor(xor(IN48, IN2), IN5)))) & ((xor(xor(IN45 & IN7, IN16 | IN6), IN37)) & ((!(IN35)) | (!(IN34))))) & (IN30 & ((!(IN5 | IN39)) & IN24))) & ((xor(xor(false, xor(xor(IN9, (IN26 | IN23) | (IN11 | IN43)), !(xor(xor(IN43, IN8), IN5)))), xor(xor(IN14, !(IN40 & IN5)), (IN6 | IN9) & (!(IN19))))) | (!(!((IN32 | IN42) | (!(IN2))))))) | (!((!(xor(xor(xor(xor(IN8 & IN44, !(IN27)), IN30 & IN14), xor(xor(xor(xor(true, IN38), IN6), IN42 & IN45), IN38 | IN48)), xor(xor(IN40, !(IN38)), IN43 | IN46)))) & (xor(xor(!(IN3), xor(xor(false & (IN3 & IN19), IN18), !(IN9 & IN41))), ((IN34 | IN41) & IN25) | (IN17 & (xor(xor(IN11, IN5), IN40)))))))), ((!(xor(xor(IN12, !(!(IN45 | IN38))), (xor(xor(IN8 & IN43, IN16 | IN4), IN18)) & ((xor(xor(IN2, IN13), IN22)) & IN38)))) & ((xor(xor(((xor(xor(IN34, IN30), IN44)) & (IN45 | IN14)) | IN49, (xor(xor(xor(xor(IN16, IN35), IN22), IN36 | IN17), xor(xor(IN26, IN21), IN2))) & (xor(xor(!(IN2), IN48), xor(xor(false, IN38), IN6)))), (!(IN21 & true)) & ((!(IN24)) & IN36))) & ((!(xor(xor(!(IN42), IN29 | IN47), IN31 & IN8))) & ((xor(xor(xor(xor(IN26, IN10), IN18), IN10 | IN2), IN38 & IN29)) & IN25)))) | IN7), ((xor(xor((!((!(!(IN41))) | IN27)) & ((((!(IN9)) & IN6) & (IN27 | IN6)) & (xor(xor(IN40, IN44), IN44))), IN47 & IN33), (IN42 & (((IN4 & IN43) & (IN21 & IN33)) | ((!(IN14)) | (xor(xor(IN12, IN35), IN7))))) | (xor(xor(!(IN20 & (IN21 & IN14)), xor(xor(!(IN47), !(IN35 | IN50)), xor(xor(IN12 & IN50, IN5 | IN12), IN33 | IN20))), !(xor(xor(!(IN8), IN6), !(IN23))))))) | (((IN44 | (!((IN1 | IN25) | (!(IN27))))) & ((((xor(xor(IN14, IN9), IN13)) | (xor(xor(IN36, IN37), IN40))) & (xor(xor(IN23, IN49 | IN3), IN37))) | (IN25 & ((IN1 | IN28) | (!(IN25)))))) & (!(((xor(xor(IN26 & false, xor(xor(IN13, IN29), IN15)), !(IN29))) & ((IN41 & IN7) & (IN36 & IN7))) & ((xor(xor(IN8 & IN8, IN29 & IN13), IN9 | IN26)) & (xor(xor(IN22 | IN40, IN37 | IN31), IN25 & IN44))))))) | ((!(xor(xor(!(IN43), (((!(IN44)) & (xor(xor(IN38, IN39), IN24))) & ((xor(xor(IN15, IN31), IN17)) | (xor(xor(IN44, IN39), IN24)))) | (!(IN23 | (xor(xor(IN46, IN33), IN26))))), IN49 & IN14))) | IN13)), xor(xor((((xor(xor(IN45 | (!(IN34)), !((IN22 & IN36) & (xor(xor(IN10, IN13), IN8)))), ((xor(xor(IN2, IN43), IN23)) | (xor(xor(IN41, IN20), IN3))) | (!(IN42)))) | (xor(xor(!(IN22 & (IN15 | IN36)), ((IN20 | IN29) | (IN13 & IN26)) & (!(IN2 | IN1))), !(xor(xor(IN45 | IN20, xor(xor(IN16, IN44), IN14)), IN16 | IN7))))) | ((((!(IN8)) & (IN24 & (!(IN17)))) & (((IN44 & IN23) | (IN30 | IN28)) & true)) & ((!((IN36 & IN33) | (xor(xor(IN1, IN44), IN38)))) | (IN32 & ((xor(xor(IN23, IN29), IN27)) | (!(IN49))))))) & (((xor(xor(xor(xor(!(IN9), IN1), (!(IN43)) & (xor(xor(IN14, IN27), IN30))), !(IN16)), (xor(xor(IN33 & IN28, IN19), IN24 & IN23)) & ((!(IN23)) & (IN42 & IN5)))) | ((!(xor(xor(xor(xor(IN17, IN45), IN41), !(IN5)), IN45 | IN7))) & (xor(xor(!(IN43 & IN44), !(IN1)), !(xor(xor(IN41, IN28), IN40)))))) | ((IN38 & ((!(xor(xor(IN21, IN30), IN38))) | ((IN8 & IN28) & (IN1 & true)))) | (IN39 & IN32))), (xor(xor((xor(xor(!(xor(xor(IN32 | IN37, xor(xor(IN13, IN49), IN42)), IN46)), IN13), !(!(IN50 | IN35)))) | (!(xor(xor((IN21 & IN6) & (xor(xor(IN36, IN3), IN26)), !(IN23)), (xor(xor(IN42, IN9), IN40)) & (!(IN28))))), ((!(xor(xor(IN11 & IN7, IN50), xor(xor(IN8, IN21), IN15)))) & ((xor(xor(xor(xor(IN1, IN47), IN39), xor(xor(IN32, IN41), IN50)), IN20 | IN22)) | (xor(xor(xor(xor(IN15, IN20), IN33), IN14 | IN22), IN44)))) | (((xor(xor(IN33 & IN32, IN31 & IN4), xor(xor(IN10, IN18), IN10))) & (xor(xor(!(IN46), IN38 & IN43), xor(xor(IN12, IN26), IN5)))) & IN45)), ((xor(xor((IN10 | IN16) & (xor(xor(IN43, IN14), IN48)), (xor(true, IN25)) & IN37), !(IN41 | IN29))) | (xor(xor(xor(xor(xor(xor(IN18, true), IN5), xor(xor(IN42, IN7), IN3)), !(IN8)), IN37 | (xor(xor(IN40, IN9), IN47))), !(!(IN20))))) | IN33)) | ((!(((!(IN17 & IN5)) | (IN19 | (IN21 | IN31))) & (xor(xor(IN5, !(IN19)), false)))) | IN30)), !(xor(xor((xor(xor(!(!(!(IN11))), !((IN10 & IN1) & (IN4 & IN26))), (xor(xor(IN23, !(IN47)), !(IN46))) & ((IN17 | IN33) & (IN17 | IN42)))) | (xor(xor((IN14 | IN14) & ((IN50 | IN39) | (xor(xor(IN5, IN13), IN31))), IN18), ((IN30 | IN1) | (IN17 | IN4)) | IN17)), !((xor(xor((!(IN39)) & IN28, (IN26 & IN24) | IN5), (!(IN5)) & (IN29 | IN47))) | IN17)), IN31 | ((((IN30 | IN37) | (IN49 & IN2)) & IN20) & ((!(!(IN46))) | true)))))))

*)

FUNCTION_BLOCK F_CollectInput
  VAR_IN_OUT
      Data : ARRAY[1..50] OF BOOL;
  END_VAR
  VAR_INPUT
      TICK  : BOOL := 0;
      IN1   : BOOL := 0;
      IN2   : BOOL := 0;
      IN3   : BOOL := 0;
      IN4   : BOOL := 0;
      IN5   : BOOL := 0;
      RESET : BOOL := FALSE;
  END_VAR
  VAR_OUTPUT
      Finished : BOOL;
  END_VAR
  VAR
      j    : USINT := 1;
      tock : BOOL  := 0;
  END_VAR
  IF NOT RESET AND tock = NOT TICK THEN
      Data[j]   := IN1;
      Data[j+1] := IN2;
      Data[j+2] := IN3;
      Data[j+3] := IN4;
      Data[j+4] := IN5;
      j := j + 5;
      tock := TICK;
  ELSE
      j := 1;
      tock := 0;
  END_IF;
  Finished := (j > 50);
END_FUNCTION_BLOCK

PROGRAM Boiler
  VAR
    Data  : ARRAY[1..50] OF BOOL;
    Ready : BOOL;
    CollectInput : F_CollectInput;
  END_VAR
  VAR
    TICK     AT %IX1.0 : BOOL;
    IN1      AT %IX0.3 : BOOL;
    IN2      AT %IX0.4 : BOOL;
    IN3      AT %IX0.5 : BOOL;
    IN4      AT %IX0.6 : BOOL;
    IN5      AT %IX0.7 : BOOL;
    OutReady AT %QX0.0 : BOOL := FALSE;
    FeedNext AT %QX0.1 : BOOL := FALSE;
    Out      AT %QX0.2 : BOOL;
  END_VAR
  CollectInput(TICK:=TICK, IN1:=IN1, IN2:=IN2, IN3:=IN3, IN4:=IN4, IN5:=IN5);
  Ready := CollectInput.Finished;
  FeedNext := 1;
  IF Ready THEN
    Out := ((((NOT Data[49]) XOR Data[20]) XOR (NOT (NOT ((NOT (NOT Data[20])) OR ((NOT (((Data[1] OR Data[21]) AND ((Data[13] XOR Data[2]) XOR Data[39])) AND (NOT (Data[34] OR Data[7])))) AND (NOT (NOT (((Data[4] AND Data[42]) XOR ((Data[12] XOR Data[33]) XOR Data[1])) XOR (NOT Data[24]))))))))) OR (((((((((((NOT (NOT (Data[2] AND Data[8]))) XOR (((Data[41] AND Data[1]) AND (Data[10] OR Data[13])) AND Data[47])) XOR (NOT (((Data[42] XOR Data[37]) XOR Data[36]) AND Data[20]))) AND TRUE) OR Data[48]) XOR Data[37]) XOR ((NOT ((NOT (((Data[26] XOR Data[18]) XOR Data[46]) OR (Data[49] AND Data[34]))) OR ((((Data[3] XOR Data[49]) XOR Data[16]) OR (NOT Data[33])) OR Data[21]))) AND ((((NOT (((FALSE OR Data[24]) XOR (NOT Data[1])) XOR ((Data[46] XOR Data[37]) XOR Data[21]))) AND (NOT Data[49])) XOR Data[13]) XOR (NOT ((((Data[41] OR Data[32]) OR Data[21]) XOR (((Data[18] XOR Data[1]) XOR Data[35]) OR ((Data[21] XOR Data[7]) XOR Data[35]))) XOR ((NOT Data[41]) AND (Data[27] AND Data[20]))))))) XOR ((((((Data[50] AND ((Data[19] XOR Data[26]) XOR Data[19])) AND ((NOT Data[47]) AND ((Data[48] XOR Data[2]) XOR Data[5]))) AND ((((Data[45] AND Data[7]) XOR (Data[16] OR Data[6])) XOR Data[37]) AND ((NOT Data[35]) OR (NOT Data[34])))) AND (Data[30] AND ((NOT (Data[5] OR Data[39])) AND Data[24]))) AND (((FALSE XOR ((Data[9] XOR ((Data[26] OR Data[23]) OR (Data[11] OR Data[43]))) XOR (NOT ((Data[43] XOR Data[8]) XOR Data[5])))) XOR ((Data[14] XOR (NOT (Data[40] AND Data[5]))) XOR ((Data[6] OR Data[9]) AND (NOT Data[19])))) OR (NOT (NOT ((Data[32] OR Data[42]) OR (NOT Data[2])))))) OR (NOT ((NOT (((((Data[8] AND Data[44]) XOR (NOT Data[27])) XOR (Data[30] AND Data[14])) XOR ((((TRUE XOR Data[38]) XOR Data[6]) XOR (Data[42] AND Data[45])) XOR (Data[38] OR Data[48]))) XOR ((Data[40] XOR (NOT Data[38])) XOR (Data[43] OR Data[46])))) AND (((NOT Data[3]) XOR (((FALSE AND (Data[3] AND Data[19])) XOR Data[18]) XOR (NOT (Data[9] AND Data[41])))) XOR (((Data[34] OR Data[41]) AND Data[25]) OR (Data[17] AND ((Data[11] XOR Data[5]) XOR Data[40])))))))) XOR (((NOT ((Data[12] XOR (NOT (NOT (Data[45] OR Data[38])))) XOR ((((Data[8] AND Data[43]) XOR (Data[16] OR Data[4])) XOR Data[18]) AND (((Data[2] XOR Data[13]) XOR Data[22]) AND Data[38])))) AND (((((((Data[34] XOR Data[30]) XOR Data[44]) AND (Data[45] OR Data[14])) OR Data[49]) XOR (((((Data[16] XOR Data[35]) XOR Data[22]) XOR (Data[36] OR Data[17])) XOR ((Data[26] XOR Data[21]) XOR Data[2])) AND (((NOT Data[2]) XOR Data[48]) XOR ((FALSE XOR Data[38]) XOR Data[6])))) XOR ((NOT (Data[21] AND TRUE)) AND ((NOT Data[24]) AND Data[36]))) AND ((NOT (((NOT Data[42]) XOR (Data[29] OR Data[47])) XOR (Data[31] AND Data[8]))) AND (((((Data[26] XOR Data[10]) XOR Data[18]) XOR (Data[10] OR Data[2])) XOR (Data[38] AND Data[29])) AND Data[25])))) OR Data[7])) XOR ((((((NOT ((NOT (NOT Data[41])) OR Data[27])) AND ((((NOT Data[9]) AND Data[6]) AND (Data[27] OR Data[6])) AND ((Data[40] XOR Data[44]) XOR Data[44]))) XOR (Data[47] AND Data[33])) XOR ((Data[42] AND (((Data[4] AND Data[43]) AND (Data[21] AND Data[33])) OR ((NOT Data[14]) OR ((Data[12] XOR Data[35]) XOR Data[7])))) OR (((NOT (Data[20] AND (Data[21] AND Data[14]))) XOR (((NOT Data[47]) XOR (NOT (Data[35] OR Data[50]))) XOR (((Data[12] AND Data[50]) XOR (Data[5] OR Data[12])) XOR (Data[33] OR Data[20])))) XOR (NOT (((NOT Data[8]) XOR Data[6]) XOR (NOT Data[23])))))) OR (((Data[44] OR (NOT ((Data[1] OR Data[25]) OR (NOT Data[27])))) AND (((((Data[14] XOR Data[9]) XOR Data[13]) OR ((Data[36] XOR Data[37]) XOR Data[40])) AND ((Data[23] XOR (Data[49] OR Data[3])) XOR Data[37])) OR (Data[25] AND ((Data[1] OR Data[28]) OR (NOT Data[25]))))) AND (NOT (((((Data[26] AND FALSE) XOR ((Data[13] XOR Data[29]) XOR Data[15])) XOR (NOT Data[29])) AND ((Data[41] AND Data[7]) AND (Data[36] AND Data[7]))) AND ((((Data[8] AND Data[8]) XOR (Data[29] AND Data[13])) XOR (Data[9] OR Data[26])) AND (((Data[22] OR Data[40]) XOR (Data[37] OR Data[31])) XOR (Data[25] AND Data[44]))))))) OR ((NOT (((NOT Data[43]) XOR ((((NOT Data[44]) AND ((Data[38] XOR Data[39]) XOR Data[24])) AND (((Data[15] XOR Data[31]) XOR Data[17]) OR ((Data[44] XOR Data[39]) XOR Data[24]))) OR (NOT (Data[23] OR ((Data[46] XOR Data[33]) XOR Data[26]))))) XOR (Data[49] AND Data[14]))) OR Data[13]))) XOR ((((((((Data[45] OR (NOT Data[34])) XOR (NOT ((Data[22] AND Data[36]) AND ((Data[10] XOR Data[13]) XOR Data[8])))) XOR ((((Data[2] XOR Data[43]) XOR Data[23]) OR ((Data[41] XOR Data[20]) XOR Data[3])) OR (NOT Data[42]))) OR (((NOT (Data[22] AND (Data[15] OR Data[36]))) XOR (((Data[20] OR Data[29]) OR (Data[13] AND Data[26])) AND (NOT (Data[2] OR Data[1])))) XOR (NOT (((Data[45] OR Data[20]) XOR ((Data[16] XOR Data[44]) XOR Data[14])) XOR (Data[16] OR Data[7]))))) OR ((((NOT Data[8]) AND (Data[24] AND (NOT Data[17]))) AND (((Data[44] AND Data[23]) OR (Data[30] OR Data[28])) AND TRUE)) AND ((NOT ((Data[36] AND Data[33]) OR ((Data[1] XOR Data[44]) XOR Data[38]))) OR (Data[32] AND (((Data[23] XOR Data[29]) XOR Data[27]) OR (NOT Data[49])))))) AND (((((((NOT Data[9]) XOR Data[1]) XOR ((NOT Data[43]) AND ((Data[14] XOR Data[27]) XOR Data[30]))) XOR (NOT Data[16])) XOR ((((Data[33] AND Data[28]) XOR Data[19]) XOR (Data[24] AND Data[23])) AND ((NOT Data[23]) AND (Data[42] AND Data[5])))) OR ((NOT ((((Data[17] XOR Data[45]) XOR Data[41]) XOR (NOT Data[5])) XOR (Data[45] OR Data[7]))) AND (((NOT (Data[43] AND Data[44])) XOR (NOT Data[1])) XOR (NOT ((Data[41] XOR Data[28]) XOR Data[40]))))) OR ((Data[38] AND ((NOT ((Data[21] XOR Data[30]) XOR Data[38])) OR ((Data[8] AND Data[28]) AND (Data[1] AND TRUE)))) OR (Data[39] AND Data[32])))) XOR (((((((NOT (((Data[32] OR Data[37]) XOR ((Data[13] XOR Data[49]) XOR Data[42])) XOR Data[46])) XOR Data[13]) XOR (NOT (NOT (Data[50] OR Data[35])))) OR (NOT ((((Data[21] AND Data[6]) AND ((Data[36] XOR Data[3]) XOR Data[26])) XOR (NOT Data[23])) XOR (((Data[42] XOR Data[9]) XOR Data[40]) AND (NOT Data[28]))))) XOR (((NOT (((Data[11] AND Data[7]) XOR Data[50]) XOR ((Data[8] XOR Data[21]) XOR Data[15]))) AND (((((Data[1] XOR Data[47]) XOR Data[39]) XOR ((Data[32] XOR Data[41]) XOR Data[50])) XOR (Data[20] OR Data[22])) OR ((((Data[15] XOR Data[20]) XOR Data[33]) XOR (Data[14] OR Data[22])) XOR Data[44]))) OR (((((Data[33] AND Data[32]) XOR (Data[31] AND Data[4])) XOR ((Data[10] XOR Data[18]) XOR Data[10])) AND (((NOT Data[46]) XOR (Data[38] AND Data[43])) XOR ((Data[12] XOR Data[26]) XOR Data[5]))) AND Data[45]))) XOR ((((((Data[10] OR Data[16]) AND ((Data[43] XOR Data[14]) XOR Data[48])) XOR ((TRUE XOR Data[25]) AND Data[37])) XOR (NOT (Data[41] OR Data[29]))) OR ((((((Data[18] XOR TRUE) XOR Data[5]) XOR ((Data[42] XOR Data[7]) XOR Data[3])) XOR (NOT Data[8])) XOR (Data[37] OR ((Data[40] XOR Data[9]) XOR Data[47]))) XOR (NOT (NOT Data[20])))) OR Data[33])) OR ((NOT (((NOT (Data[17] AND Data[5])) OR (Data[19] OR (Data[21] OR Data[31]))) AND ((Data[5] XOR (NOT Data[19])) XOR FALSE))) OR Data[30]))) XOR (NOT ((((((NOT (NOT (NOT Data[11]))) XOR (NOT ((Data[10] AND Data[1]) AND (Data[4] AND Data[26])))) XOR (((Data[23] XOR (NOT Data[47])) XOR (NOT Data[46])) AND ((Data[17] OR Data[33]) AND (Data[17] OR Data[42])))) OR ((((Data[14] OR Data[14]) AND ((Data[50] OR Data[39]) OR ((Data[5] XOR Data[13]) XOR Data[31]))) XOR Data[18]) XOR (((Data[30] OR Data[1]) OR (Data[17] OR Data[4])) OR Data[17]))) XOR (NOT (((((NOT Data[39]) AND Data[28]) XOR ((Data[26] AND Data[24]) OR Data[5])) XOR ((NOT Data[5]) AND (Data[29] OR Data[47]))) OR Data[17]))) XOR (Data[31] OR ((((Data[30] OR Data[37]) OR (Data[49] AND Data[2])) AND Data[20]) AND ((NOT (NOT Data[46])) OR TRUE))))))));
    OutReady := 1;
    CollectInput(RESET:=TRUE);
  END_IF;
END_PROGRAM

CONFIGURATION Config0
  RESOURCE Res0 ON PLC
    TASK task0(INTERVAL := T#20ms,PRIORITY := 0);
    PROGRAM instance0 WITH task0 : Boiler;
  END_RESOURCE
END_CONFIGURATION
